  movel([-0.121105, -0.793361, -2.803748, -1.115280, 1.570796, 1.449692],accel_mss,speed_ms,0,blend_radius_m)
  movel([-0.120159, -0.793542, -2.803719, -1.115129, 1.570796, 1.450637],accel_mss,speed_ms,0,blend_radius_m)
  movel([-0.119008, -0.795086, -2.803467, -1.113836, 1.570796, 1.451789],accel_mss,speed_ms,0,blend_radius_m)
  movel([-0.118135, -0.797911, -2.803003, -1.111475, 1.570796, 1.452661],accel_mss,speed_ms,0,blend_radius_m)
  movel([-0.117601, -0.801037, -2.802486, -1.108866, 1.570796, 1.453195],accel_mss,speed_ms,0,blend_radius_m)
  movel([-0.115239, -0.796332, -2.803263, -1.112794, 1.570796, 1.455558],accel_mss,speed_ms,0,blend_radius_m)
  movel([-0.112520, -0.791566, -2.804039, -1.116785, 1.570796, 1.458276],accel_mss,speed_ms,0,blend_radius_m)
  movel([-0.109499, -0.786802, -2.804803, -1.120785, 1.570796, 1.461298],accel_mss,speed_ms,0,blend_radius_m)
  movel([-0.106241, -0.782109, -2.805544, -1.124735, 1.570796, 1.464556],accel_mss,speed_ms,0,blend_radius_m)
  movel([-0.099689, -0.772678, -2.807001, -1.132710, 1.570796, 1.471108],accel_mss,speed_ms,0,blend_radius_m)
  movel([-0.097728, -0.770078, -2.807395, -1.134915, 1.570796, 1.473068],accel_mss,speed_ms,0,blend_radius_m)
  movel([-0.095794, -0.767754, -2.807745, -1.136890, 1.570796, 1.475003],accel_mss,speed_ms,0,blend_radius_m)
  movel([-0.093954, -0.765885, -2.808024, -1.138480, 1.570796, 1.476842],accel_mss,speed_ms,0,blend_radius_m)
  movel([-0.092299, -0.764660, -2.808206, -1.139523, 1.570796, 1.478498],accel_mss,speed_ms,0,blend_radius_m)
  movel([-0.090884, -0.764292, -2.808260, -1.139836, 1.570796, 1.479912],accel_mss,speed_ms,0,blend_radius_m)
  movel([-0.089878, -0.764818, -2.808182, -1.139389, 1.570796, 1.480919],accel_mss,speed_ms,0,blend_radius_m)
  movel([-0.089251, -0.766042, -2.808000, -1.138346, 1.570796, 1.481545],accel_mss,speed_ms,0,blend_radius_m)
  movel([-0.088991, -0.767774, -2.807742, -1.136873, 1.570796, 1.481805],accel_mss,speed_ms,0,blend_radius_m)
  movel([-0.089073, -0.769817, -2.807435, -1.135137, 1.570796, 1.481724],accel_mss,speed_ms,0,blend_radius_m)
  movel([-0.089471, -0.771972, -2.807109, -1.133309, 1.570796, 1.481326],accel_mss,speed_ms,0,blend_radius_m)
  movel([-0.090165, -0.774050, -2.806792, -1.131547, 1.570796, 1.480631],accel_mss,speed_ms,0,blend_radius_m)
  movel([-0.091138, -0.775860, -2.806515, -1.130015, 1.570796, 1.479658],accel_mss,speed_ms,0,blend_radius_m)
  movel([-0.085055, -0.767504, -2.807782, -1.137103, 1.570796, 1.485742],accel_mss,speed_ms,0,blend_radius_m)
  movel([-0.081792, -0.763433, -2.808387, -1.140568, 1.570796, 1.489004],accel_mss,speed_ms,0,blend_radius_m)
  movel([-0.078396, -0.759483, -2.808967, -1.143939, 1.570796, 1.492400],accel_mss,speed_ms,0,blend_radius_m)
  movel([-0.074888, -0.755690, -2.809517, -1.147182, 1.570796, 1.495909],accel_mss,speed_ms,0,blend_radius_m)
  movel([-0.071275, -0.752094, -2.810031, -1.150264, 1.570796, 1.499521],accel_mss,speed_ms,0,blend_radius_m)
  movel([-0.067576, -0.748733, -2.810507, -1.153150, 1.570796, 1.503221],accel_mss,speed_ms,0,blend_radius_m)
  movel([-0.063806, -0.745643, -2.810939, -1.155807, 1.570796, 1.506991],accel_mss,speed_ms,0,blend_radius_m)
  movel([-0.061242, -0.744068, -2.811158, -1.157163, 1.570796, 1.509554],accel_mss,speed_ms,0,blend_radius_m)
  movel([-0.058496, -0.743084, -2.811294, -1.158011, 1.570796, 1.512301],accel_mss,speed_ms,0,blend_radius_m)
  movel([-0.057304, -0.742971, -2.811309, -1.158108, 1.570796, 1.513493],accel_mss,speed_ms,0,blend_radius_m)
  movel([-0.056360, -0.743186, -2.811280, -1.157923, 1.570796, 1.514437],accel_mss,speed_ms,0,blend_radius_m)
  movel([-0.055759, -0.743792, -2.811196, -1.157401, 1.570796, 1.515037],accel_mss,speed_ms,0,blend_radius_m)
  movel([-0.055607, -0.744852, -2.811049, -1.156488, 1.570796, 1.515190],accel_mss,speed_ms,0,blend_radius_m)
  movel([-0.055970, -0.746235, -2.810857, -1.155298, 1.570796, 1.514827],accel_mss,speed_ms,0,blend_radius_m)
  movel([-0.056714, -0.747783, -2.810640, -1.153965, 1.570796, 1.514083],accel_mss,speed_ms,0,blend_radius_m)
  movel([-0.058927, -0.751255, -2.810150, -1.150983, 1.570796, 1.511869],accel_mss,speed_ms,0,blend_radius_m)
  movel([-0.061573, -0.754500, -2.809688, -1.148201, 1.570796, 1.509223],accel_mss,speed_ms,0,blend_radius_m)
  movel([-0.064470, -0.757491, -2.809257, -1.145642, 1.570796, 1.506326],accel_mss,speed_ms,0,blend_radius_m)
  movel([-0.067437, -0.760200, -2.808862, -1.143327, 1.570796, 1.503359],accel_mss,speed_ms,0,blend_radius_m)
  movel([-0.063607, -0.758678, -2.809084, -1.144626, 1.570796, 1.507189],accel_mss,speed_ms,0,blend_radius_m)
  movel([-0.059620, -0.756697, -2.809371, -1.146320, 1.570796, 1.511176],accel_mss,speed_ms,0,blend_radius_m)
  movel([-0.055519, -0.754282, -2.809719, -1.148388, 1.570796, 1.515278],accel_mss,speed_ms,0,blend_radius_m)
  movel([-0.051338, -0.751454, -2.810122, -1.150813, 1.570796, 1.519459],accel_mss,speed_ms,0,blend_radius_m)
  movel([-0.048030, -0.748869, -2.810488, -1.153033, 1.570796, 1.522766],accel_mss,speed_ms,0,blend_radius_m)
  movel([-0.041537, -0.743272, -2.811268, -1.157849, 1.570796, 1.529259],accel_mss,speed_ms,0,blend_radius_m)
  movel([-0.038202, -0.740640, -2.811630, -1.160119, 1.570796, 1.532595],accel_mss,speed_ms,0,blend_radius_m)
  movel([-0.034400, -0.737919, -2.812001, -1.162470, 1.570796, 1.536396],accel_mss,speed_ms,0,blend_radius_m)
  movel([-0.027997, -0.733681, -2.812571, -1.166137, 1.570796, 1.542799],accel_mss,speed_ms,0,blend_radius_m)
  movel([-0.024935, -0.731926, -2.812805, -1.167658, 1.570796, 1.545861],accel_mss,speed_ms,0,blend_radius_m)
  movel([-0.022568, -0.730917, -2.812939, -1.168533, 1.570796, 1.548229],accel_mss,speed_ms,0,blend_radius_m)
  movel([-0.021784, -0.730807, -2.812954, -1.168629, 1.570796, 1.549013],accel_mss,speed_ms,0,blend_radius_m)
  movel([-0.021347, -0.731026, -2.812924, -1.168438, 1.570796, 1.549449],accel_mss,speed_ms,0,blend_radius_m)
  movel([-0.021306, -0.731611, -2.812847, -1.167931, 1.570796, 1.549490],accel_mss,speed_ms,0,blend_radius_m)
  movel([-0.021722, -0.732612, -2.812714, -1.167063, 1.570796, 1.549074],accel_mss,speed_ms,0,blend_radius_m)
  movel([-0.023301, -0.735118, -2.812379, -1.164892, 1.570796, 1.547495],accel_mss,speed_ms,0,blend_radius_m)
  movel([-0.025347, -0.737745, -2.812024, -1.162620, 1.570796, 1.545450],accel_mss,speed_ms,0,blend_radius_m)
  movel([-0.027725, -0.740428, -2.811659, -1.160302, 1.570796, 1.543072],accel_mss,speed_ms,0,blend_radius_m)
  movel([-0.030292, -0.743084, -2.811294, -1.158011, 1.570796, 1.540504],accel_mss,speed_ms,0,blend_radius_m)
  movel([-0.035478, -0.748036, -2.810605, -1.153749, 1.570796, 1.535318],accel_mss,speed_ms,0,blend_radius_m)
  movel([-0.039835, -0.752018, -2.810042, -1.150329, 1.570796, 1.530962],accel_mss,speed_ms,0,blend_radius_m)
  movel([-0.037640, -0.751618, -2.810099, -1.150672, 1.570796, 1.533156],accel_mss,speed_ms,0,blend_radius_m)
  movel([-0.035326, -0.750943, -2.810195, -1.151251, 1.570796, 1.535470],accel_mss,speed_ms,0,blend_radius_m)
  movel([-0.030418, -0.748918, -2.810481, -1.152991, 1.570796, 1.540378],accel_mss,speed_ms,0,blend_radius_m)
  movel([-0.025249, -0.746199, -2.810862, -1.155329, 1.570796, 1.545548],accel_mss,speed_ms,0,blend_radius_m)
  movel([-0.019955, -0.743049, -2.811299, -1.158041, 1.570796, 1.550841],accel_mss,speed_ms,0,blend_radius_m)
  movel([-0.015550, -0.740169, -2.811694, -1.160526, 1.570796, 1.555246],accel_mss,speed_ms,0,blend_radius_m)
  movel([-0.002182, -0.730928, -2.812937, -1.168523, 1.570796, 1.568614],accel_mss,speed_ms,0,blend_radius_m)
  movel([0.000291, -0.729638, -2.813108, -1.169643, 1.570796, 1.571087],accel_mss,speed_ms,0,blend_radius_m)
  movel([0.002219, -0.729213, -2.813164, -1.170012, 1.570796, 1.573015],accel_mss,speed_ms,0,blend_radius_m)
  movel([0.002614, -0.729532, -2.813122, -1.169735, 1.570796, 1.573410],accel_mss,speed_ms,0,blend_radius_m)
  movel([0.002432, -0.730316, -2.813018, -1.169054, 1.570796, 1.573228],accel_mss,speed_ms,0,blend_radius_m)
  movel([0.001528, -0.731648, -2.812842, -1.167899, 1.570796, 1.572325],accel_mss,speed_ms,0,blend_radius_m)
  movel([-0.000242, -0.733605, -2.812581, -1.166203, 1.570796, 1.570554],accel_mss,speed_ms,0,blend_radius_m)
  movel([-0.003204, -0.736443, -2.812200, -1.163745, 1.570796, 1.567592],accel_mss,speed_ms,0,blend_radius_m)
  movel([-0.006618, -0.739358, -2.811805, -1.161226, 1.570796, 1.564179],accel_mss,speed_ms,0,blend_radius_m)
  movel([-0.009977, -0.741812, -2.811469, -1.159108, 1.570796, 1.560819],accel_mss,speed_ms,0,blend_radius_m)
  movel([-0.011482, -0.742703, -2.811346, -1.158339, 1.570796, 1.559315],accel_mss,speed_ms,0,blend_radius_m)
  movel([-0.012779, -0.743271, -2.811268, -1.157850, 1.570796, 1.558017],accel_mss,speed_ms,0,blend_radius_m)
  movel([-0.007737, -0.743073, -2.811295, -1.158021, 1.570796, 1.563059],accel_mss,speed_ms,0,blend_radius_m)
  movel([-0.002332, -0.742171, -2.811420, -1.158799, 1.570796, 1.568464],accel_mss,speed_ms,0,blend_radius_m)
  movel([0.003362, -0.740698, -2.811622, -1.160069, 1.570796, 1.574158],accel_mss,speed_ms,0,blend_radius_m)
  movel([0.009278, -0.738793, -2.811882, -1.161714, 1.570796, 1.580074],accel_mss,speed_ms,0,blend_radius_m)
  movel([0.021466, -0.734216, -2.812500, -1.165673, 1.570796, 1.592262],accel_mss,speed_ms,0,blend_radius_m)
  movel([0.033600, -0.729546, -2.813120, -1.169723, 1.570796, 1.604396],accel_mss,speed_ms,0,blend_radius_m)
  movel([0.035605, -0.729117, -2.813177, -1.170096, 1.570796, 1.606402],accel_mss,speed_ms,0,blend_radius_m)
  movel([0.036255, -0.729398, -2.813140, -1.169851, 1.570796, 1.607051],accel_mss,speed_ms,0,blend_radius_m)
  movel([0.036422, -0.730219, -2.813031, -1.169139, 1.570796, 1.607218],accel_mss,speed_ms,0,blend_radius_m)
  movel([0.036036, -0.731427, -2.812871, -1.168090, 1.570796, 1.606833],accel_mss,speed_ms,0,blend_radius_m)
  movel([0.034004, -0.734771, -2.812425, -1.165193, 1.570796, 1.604800],accel_mss,speed_ms,0,blend_radius_m)
  movel([0.032557, -0.736690, -2.812167, -1.163532, 1.570796, 1.603354],accel_mss,speed_ms,0,blend_radius_m)
  movel([0.029315, -0.740256, -2.811682, -1.160451, 1.570796, 1.600111],accel_mss,speed_ms,0,blend_radius_m)
  movel([0.025758, -0.743429, -2.811246, -1.157714, 1.570796, 1.596555],accel_mss,speed_ms,0,blend_radius_m)
  movel([0.022037, -0.746209, -2.810860, -1.155320, 1.570796, 1.592834],accel_mss,speed_ms,0,blend_radius_m)
  movel([0.018315, -0.748574, -2.810529, -1.153286, 1.570796, 1.589112],accel_mss,speed_ms,0,blend_radius_m)
  movel([0.014745, -0.750516, -2.810255, -1.151618, 1.570796, 1.585541],accel_mss,speed_ms,0,blend_radius_m)
  movel([0.011481, -0.752014, -2.810043, -1.150332, 1.570796, 1.582277],accel_mss,speed_ms,0,blend_radius_m)
  movel([0.008687, -0.753044, -2.809896, -1.149449, 1.570796, 1.579483],accel_mss,speed_ms,0,blend_radius_m)
  movel([0.008653, -0.753899, -2.809774, -1.148717, 1.570796, 1.579449],accel_mss,speed_ms,0,blend_radius_m)
  movel([0.009139, -0.754307, -2.809715, -1.148367, 1.570796, 1.579935],accel_mss,speed_ms,0,blend_radius_m)
  movel([0.010647, -0.754705, -2.809658, -1.148026, 1.570796, 1.581444],accel_mss,speed_ms,0,blend_radius_m)
  movel([0.012360, -0.754771, -2.809649, -1.147969, 1.570796, 1.583157],accel_mss,speed_ms,0,blend_radius_m)
  movel([0.016128, -0.754316, -2.809714, -1.148359, 1.570796, 1.586925],accel_mss,speed_ms,0,blend_radius_m)
  movel([0.022850, -0.753072, -2.809892, -1.149425, 1.570796, 1.593647],accel_mss,speed_ms,0,blend_radius_m)
  movel([0.029687, -0.751537, -2.810110, -1.150742, 1.570796, 1.600483],accel_mss,speed_ms,0,blend_radius_m)
  movel([0.043712, -0.747708, -2.810651, -1.154030, 1.570796, 1.614508],accel_mss,speed_ms,0,blend_radius_m)
  movel([0.047601, -0.746731, -2.810787, -1.154870, 1.570796, 1.618397],accel_mss,speed_ms,0,blend_radius_m)
  movel([0.050057, -0.746348, -2.810841, -1.155200, 1.570796, 1.620854],accel_mss,speed_ms,0,blend_radius_m)
  movel([0.052405, -0.746275, -2.810851, -1.155263, 1.570796, 1.623201],accel_mss,speed_ms,0,blend_radius_m)
  movel([0.054288, -0.746698, -2.810792, -1.154899, 1.570796, 1.625084],accel_mss,speed_ms,0,blend_radius_m)
  movel([0.055366, -0.747783, -2.810640, -1.153965, 1.570796, 1.626162],accel_mss,speed_ms,0,blend_radius_m)
  movel([0.055503, -0.748623, -2.810522, -1.153244, 1.570796, 1.626300],accel_mss,speed_ms,0,blend_radius_m)
  movel([0.055317, -0.749691, -2.810372, -1.152326, 1.570796, 1.626113],accel_mss,speed_ms,0,blend_radius_m)
  movel([0.054755, -0.751016, -2.810184, -1.151188, 1.570796, 1.625552],accel_mss,speed_ms,0,blend_radius_m)
  movel([0.053791, -0.752605, -2.809958, -1.149825, 1.570796, 1.624588],accel_mss,speed_ms,0,blend_radius_m)
  movel([0.052380, -0.754061, -2.809750, -1.148578, 1.570796, 1.623176],accel_mss,speed_ms,0,blend_radius_m)
  movel([0.050460, -0.755437, -2.809553, -1.147399, 1.570796, 1.621256],accel_mss,speed_ms,0,blend_radius_m)
  movel([0.040183, -0.761646, -2.808651, -1.142093, 1.570796, 1.610979],accel_mss,speed_ms,0,blend_radius_m)
  movel([0.036738, -0.763274, -2.808411, -1.140704, 1.570796, 1.607535],accel_mss,speed_ms,0,blend_radius_m)
  movel([0.035260, -0.763727, -2.808344, -1.140318, 1.570796, 1.606056],accel_mss,speed_ms,0,blend_radius_m)
  movel([0.034042, -0.763830, -2.808329, -1.140230, 1.570796, 1.604838],accel_mss,speed_ms,0,blend_radius_m)
  movel([0.039097, -0.765388, -2.808098, -1.138903, 1.570796, 1.609893],accel_mss,speed_ms,0,blend_radius_m)
  movel([0.044720, -0.766036, -2.808001, -1.138351, 1.570796, 1.615516],accel_mss,speed_ms,0,blend_radius_m)
  movel([0.050778, -0.765942, -2.808015, -1.138432, 1.570796, 1.621574],accel_mss,speed_ms,0,blend_radius_m)
  movel([0.057144, -0.765260, -2.808117, -1.139012, 1.570796, 1.627940],accel_mss,speed_ms,0,blend_radius_m)
  movel([0.062648, -0.763858, -2.808325, -1.140207, 1.570796, 1.633444],accel_mss,speed_ms,0,blend_radius_m)
  movel([0.070534, -0.762014, -2.808596, -1.141778, 1.570796, 1.641330],accel_mss,speed_ms,0,blend_radius_m)
  movel([0.074102, -0.761631, -2.808653, -1.142105, 1.570796, 1.644899],accel_mss,speed_ms,0,blend_radius_m)
  movel([0.076754, -0.761962, -2.808604, -1.141823, 1.570796, 1.647550],accel_mss,speed_ms,0,blend_radius_m)
  movel([0.077577, -0.762479, -2.808528, -1.141382, 1.570796, 1.648374],accel_mss,speed_ms,0,blend_radius_m)
  movel([0.077981, -0.763272, -2.808411, -1.140706, 1.570796, 1.648777],accel_mss,speed_ms,0,blend_radius_m)
  movel([0.077904, -0.764377, -2.808248, -1.139764, 1.570796, 1.648701],accel_mss,speed_ms,0,blend_radius_m)
  movel([0.077296, -0.765814, -2.808034, -1.138540, 1.570796, 1.648093],accel_mss,speed_ms,0,blend_radius_m)
  movel([0.076368, -0.767285, -2.807815, -1.137289, 1.570796, 1.647164],accel_mss,speed_ms,0,blend_radius_m)
  movel([0.075295, -0.768687, -2.807605, -1.136097, 1.570796, 1.646091],accel_mss,speed_ms,0,blend_radius_m)
  movel([0.072924, -0.771293, -2.807212, -1.133884, 1.570796, 1.643720],accel_mss,speed_ms,0,blend_radius_m)
  movel([0.070302, -0.773862, -2.806821, -1.131706, 1.570796, 1.641099],accel_mss,speed_ms,0,blend_radius_m)
  movel([0.064988, -0.778418, -2.806120, -1.127851, 1.570796, 1.635784],accel_mss,speed_ms,0,blend_radius_m)
  movel([0.062326, -0.780386, -2.805814, -1.126189, 1.570796, 1.633122],accel_mss,speed_ms,0,blend_radius_m)
  movel([0.067181, -0.779786, -2.805907, -1.126695, 1.570796, 1.637977],accel_mss,speed_ms,0,blend_radius_m)
  movel([0.072189, -0.778807, -2.806060, -1.127523, 1.570796, 1.642985],accel_mss,speed_ms,0,blend_radius_m)
  movel([0.077338, -0.777493, -2.806263, -1.128633, 1.570796, 1.648134],accel_mss,speed_ms,0,blend_radius_m)
  movel([0.082615, -0.775877, -2.806512, -1.130000, 1.570796, 1.653412],accel_mss,speed_ms,0,blend_radius_m)
  movel([0.093490, -0.771912, -2.807118, -1.133359, 1.570796, 1.664286],accel_mss,speed_ms,0,blend_radius_m)
  movel([0.104701, -0.767216, -2.807825, -1.137348, 1.570796, 1.675497],accel_mss,speed_ms,0,blend_radius_m)
  movel([0.107639, -0.766300, -2.807962, -1.138127, 1.570796, 1.678435],accel_mss,speed_ms,0,blend_radius_m)
  movel([0.108683, -0.766493, -2.807933, -1.137963, 1.570796, 1.679480],accel_mss,speed_ms,0,blend_radius_m)
  movel([0.109107, -0.767448, -2.807791, -1.137151, 1.570796, 1.679903],accel_mss,speed_ms,0,blend_radius_m)
  movel([0.108974, -0.768426, -2.807644, -1.136319, 1.570796, 1.679770],accel_mss,speed_ms,0,blend_radius_m)
  movel([0.108569, -0.769523, -2.807479, -1.135387, 1.570796, 1.679365],accel_mss,speed_ms,0,blend_radius_m)
  movel([0.107060, -0.772017, -2.807102, -1.133270, 1.570796, 1.677856],accel_mss,speed_ms,0,blend_radius_m)
  movel([0.104857, -0.774737, -2.806687, -1.130965, 1.570796, 1.675653],accel_mss,speed_ms,0,blend_radius_m)
  movel([0.102226, -0.777515, -2.806260, -1.128615, 1.570796, 1.673022],accel_mss,speed_ms,0,blend_radius_m)
  movel([0.096762, -0.782520, -2.805480, -1.124390, 1.570796, 1.667558],accel_mss,speed_ms,0,blend_radius_m)
  movel([0.092780, -0.785621, -2.804990, -1.121778, 1.570796, 1.663577],accel_mss,speed_ms,0,blend_radius_m)
  movel([0.095018, -0.784942, -2.805098, -1.122349, 1.570796, 1.665815],accel_mss,speed_ms,0,blend_radius_m)
  movel([0.097342, -0.784002, -2.805247, -1.123140, 1.570796, 1.668138],accel_mss,speed_ms,0,blend_radius_m)
  movel([0.102193, -0.781425, -2.805652, -1.125313, 1.570796, 1.672990],accel_mss,speed_ms,0,blend_radius_m)
  movel([0.107238, -0.777995, -2.806185, -1.128209, 1.570796, 1.678035],accel_mss,speed_ms,0,blend_radius_m)
  movel([0.112383, -0.773843, -2.806824, -1.131722, 1.570796, 1.683179],accel_mss,speed_ms,0,blend_radius_m)
  movel([0.117534, -0.769067, -2.807548, -1.135774, 1.570796, 1.688330],accel_mss,speed_ms,0,blend_radius_m)
  movel([0.122590, -0.763799, -2.808333, -1.140256, 1.570796, 1.693387],accel_mss,speed_ms,0,blend_radius_m)
  movel([0.127452, -0.758145, -2.809162, -1.145082, 1.570796, 1.698249],accel_mss,speed_ms,0,blend_radius_m)
  movel([0.132018, -0.752235, -2.810011, -1.150143, 1.570796, 1.702814],accel_mss,speed_ms,0,blend_radius_m)
  movel([0.134037, -0.749592, -2.810386, -1.152411, 1.570796, 1.704834],accel_mss,speed_ms,0,blend_radius_m)
  movel([0.135120, -0.748440, -2.810548, -1.153401, 1.570796, 1.705916],accel_mss,speed_ms,0,blend_radius_m)
  movel([0.136237, -0.747552, -2.810672, -1.154164, 1.570796, 1.707033],accel_mss,speed_ms,0,blend_radius_m)
  movel([0.137379, -0.747065, -2.810741, -1.154583, 1.570796, 1.708175],accel_mss,speed_ms,0,blend_radius_m)
  movel([0.138333, -0.747027, -2.810746, -1.154616, 1.570796, 1.709129],accel_mss,speed_ms,0,blend_radius_m)
  movel([0.139345, -0.747698, -2.810652, -1.154039, 1.570796, 1.710141],accel_mss,speed_ms,0,blend_radius_m)
  movel([0.139829, -0.749137, -2.810450, -1.152802, 1.570796, 1.710625],accel_mss,speed_ms,0,blend_radius_m)
  movel([0.139879, -0.751150, -2.810165, -1.151074, 1.570796, 1.710675],accel_mss,speed_ms,0,blend_radius_m)
  movel([0.139591, -0.753557, -2.809823, -1.149009, 1.570796, 1.710387],accel_mss,speed_ms,0,blend_radius_m)
  movel([0.138373, -0.758783, -2.809069, -1.144537, 1.570796, 1.709169],accel_mss,speed_ms,0,blend_radius_m)
  movel([0.136926, -0.763333, -2.808402, -1.140654, 1.570796, 1.707723],accel_mss,speed_ms,0,blend_radius_m)
  movel([0.140852, -0.757577, -2.809244, -1.145568, 1.570796, 1.711648],accel_mss,speed_ms,0,blend_radius_m)
  movel([0.144402, -0.751708, -2.810086, -1.150595, 1.570796, 1.715198],accel_mss,speed_ms,0,blend_radius_m)
  movel([0.147549, -0.745784, -2.810919, -1.155685, 1.570796, 1.718345],accel_mss,speed_ms,0,blend_radius_m)
  movel([0.150273, -0.739888, -2.811733, -1.160768, 1.570796, 1.721070],accel_mss,speed_ms,0,blend_radius_m)
  movel([0.152533, -0.734096, -2.812516, -1.165777, 1.570796, 1.723330],accel_mss,speed_ms,0,blend_radius_m)
  movel([0.154318, -0.728473, -2.813261, -1.170655, 1.570796, 1.725114],accel_mss,speed_ms,0,blend_radius_m)
  movel([0.155580, -0.723118, -2.813958, -1.175313, 1.570796, 1.726376],accel_mss,speed_ms,0,blend_radius_m)
  movel([0.156297, -0.718102, -2.814598, -1.179688, 1.570796, 1.727094],accel_mss,speed_ms,0,blend_radius_m)
  movel([0.156402, -0.711752, -2.815393, -1.185243, 1.570796, 1.727198],accel_mss,speed_ms,0,blend_radius_m)
  movel([0.156716, -0.708235, -2.815826, -1.188328, 1.570796, 1.727512],accel_mss,speed_ms,0,blend_radius_m)
  movel([0.157110, -0.706436, -2.816045, -1.189908, 1.570796, 1.727906],accel_mss,speed_ms,0,blend_radius_m)
  movel([0.157721, -0.704629, -2.816264, -1.191496, 1.570796, 1.728517],accel_mss,speed_ms,0,blend_radius_m)
  movel([0.159157, -0.701655, -2.816621, -1.194114, 1.570796, 1.729953],accel_mss,speed_ms,0,blend_radius_m)
  movel([0.160486, -0.699829, -2.816838, -1.195722, 1.570796, 1.731283],accel_mss,speed_ms,0,blend_radius_m)
  movel([0.161725, -0.698910, -2.816946, -1.196533, 1.570796, 1.732521],accel_mss,speed_ms,0,blend_radius_m)
  movel([0.162880, -0.698652, -2.816977, -1.196760, 1.570796, 1.733676],accel_mss,speed_ms,0,blend_radius_m)
  movel([0.165920, -0.699423, -2.816886, -1.196081, 1.570796, 1.736716],accel_mss,speed_ms,0,blend_radius_m)
  movel([0.166833, -0.699369, -2.816892, -1.196128, 1.570796, 1.737629],accel_mss,speed_ms,0,blend_radius_m)
  movel([0.168876, -0.694954, -2.817410, -1.200024, 1.570796, 1.739672],accel_mss,speed_ms,0,blend_radius_m)
  movel([0.170617, -0.690579, -2.817915, -1.203895, 1.570796, 1.741413],accel_mss,speed_ms,0,blend_radius_m)
  movel([0.172069, -0.686262, -2.818406, -1.207721, 1.570796, 1.742866],accel_mss,speed_ms,0,blend_radius_m)
  movel([0.173248, -0.682014, -2.818880, -1.211495, 1.570796, 1.744044],accel_mss,speed_ms,0,blend_radius_m)
  movel([0.174153, -0.677863, -2.819337, -1.215189, 1.570796, 1.744950],accel_mss,speed_ms,0,blend_radius_m)
  movel([0.174801, -0.673819, -2.819775, -1.218796, 1.570796, 1.745598],accel_mss,speed_ms,0,blend_radius_m)
  movel([0.175391, -0.666110, -2.820590, -1.225689, 1.570796, 1.746188],accel_mss,speed_ms,0,blend_radius_m)
  movel([0.175103, -0.659042, -2.821316, -1.232031, 1.570796, 1.745899],accel_mss,speed_ms,0,blend_radius_m)
  movel([0.174059, -0.652731, -2.821947, -1.237712, 1.570796, 1.744855],accel_mss,speed_ms,0,blend_radius_m)
  movel([0.172351, -0.647325, -2.822474, -1.242590, 1.570796, 1.743147],accel_mss,speed_ms,0,blend_radius_m)
  movel([0.170116, -0.642932, -2.822894, -1.246563, 1.570796, 1.740912],accel_mss,speed_ms,0,blend_radius_m)
  speed_ms = 0.005
  movel([0.170116, -0.636489, -2.816133, -1.259767, 1.570796, 1.740912],accel_mss,speed_ms,0,blend_radius_m)
  speed_ms = 0.040
  movel([0.138700, -0.661451, -2.813652, -1.237286, 1.570796, 1.709497],accel_mss,speed_ms,0,blend_radius_m)
  speed_ms = 0.005
  movel([0.138700, -0.668285, -2.820362, -1.223742, 1.570796, 1.709497],accel_mss,speed_ms,0,blend_radius_m)
  speed_ms = 0.025
  movel([0.136102, -0.667914, -2.820401, -1.224074, 1.570796, 1.706899],accel_mss,speed_ms,0,blend_radius_m)
  movel([0.133054, -0.668449, -2.820345, -1.223595, 1.570796, 1.703850],accel_mss,speed_ms,0,blend_radius_m)
  movel([0.129644, -0.669757, -2.820207, -1.222425, 1.570796, 1.700441],accel_mss,speed_ms,0,blend_radius_m)
  movel([0.125976, -0.671690, -2.820002, -1.220697, 1.570796, 1.696772],accel_mss,speed_ms,0,blend_radius_m)
  movel([0.122143, -0.674109, -2.819743, -1.218536, 1.570796, 1.692939],accel_mss,speed_ms,0,blend_radius_m)
  movel([0.118234, -0.676875, -2.819444, -1.216069, 1.570796, 1.689030],accel_mss,speed_ms,0,blend_radius_m)
  movel([0.110564, -0.682887, -2.818784, -1.210719, 1.570796, 1.681360],accel_mss,speed_ms,0,blend_radius_m)
  speed_ms = 0.005
  movel([0.110564, -0.675837, -2.812104, -1.224448, 1.570796, 1.681360],accel_mss,speed_ms,0,blend_radius_m)
  speed_ms = 0.040
  movel([0.120496, -0.667301, -2.813033, -1.232055, 1.570796, 1.691293],accel_mss,speed_ms,0,blend_radius_m)
  speed_ms = 0.005
  movel([0.120496, -0.674223, -2.819731, -1.218435, 1.570796, 1.691293],accel_mss,speed_ms,0,blend_radius_m)
  speed_ms = 0.025
  movel([0.122110, -0.669388, -2.820246, -1.222755, 1.570796, 1.692907],accel_mss,speed_ms,0,blend_radius_m)
  movel([0.123299, -0.664893, -2.820716, -1.226780, 1.570796, 1.694095],accel_mss,speed_ms,0,blend_radius_m)
  movel([0.124068, -0.660732, -2.821144, -1.230512, 1.570796, 1.694864],accel_mss,speed_ms,0,blend_radius_m)
  movel([0.124435, -0.656891, -2.821533, -1.233966, 1.570796, 1.695231],accel_mss,speed_ms,0,blend_radius_m)
  movel([0.124423, -0.653347, -2.821886, -1.237156, 1.570796, 1.695219],accel_mss,speed_ms,0,blend_radius_m)
  movel([0.124046, -0.650090, -2.822206, -1.240093, 1.570796, 1.694842],accel_mss,speed_ms,0,blend_radius_m)
  movel([0.123323, -0.647102, -2.822495, -1.242791, 1.570796, 1.694119],accel_mss,speed_ms,0,blend_radius_m)
  movel([0.122274, -0.644366, -2.822758, -1.245265, 1.570796, 1.693071],accel_mss,speed_ms,0,blend_radius_m)
  movel([0.118229, -0.637367, -2.823415, -1.251608, 1.570796, 1.689025],accel_mss,speed_ms,0,blend_radius_m)
  movel([0.116481, -0.633814, -2.823740, -1.254834, 1.570796, 1.687277],accel_mss,speed_ms,0,blend_radius_m)
  movel([0.115290, -0.629199, -2.824156, -1.259034, 1.570796, 1.686086],accel_mss,speed_ms,0,blend_radius_m)
  movel([0.114590, -0.622661, -2.824731, -1.264997, 1.570796, 1.685386],accel_mss,speed_ms,0,blend_radius_m)
  movel([0.114549, -0.615508, -2.825341, -1.271541, 1.570796, 1.685345],accel_mss,speed_ms,0,blend_radius_m)
  movel([0.115398, -0.607615, -2.825990, -1.278783, 1.570796, 1.686195],accel_mss,speed_ms,0,blend_radius_m)
  movel([0.116229, -0.603351, -2.826331, -1.282706, 1.570796, 1.687025],accel_mss,speed_ms,0,blend_radius_m)
  movel([0.117376, -0.598855, -2.826683, -1.286851, 1.570796, 1.688172],accel_mss,speed_ms,0,blend_radius_m)
  movel([0.119840, -0.591525, -2.827240, -1.293623, 1.570796, 1.690636],accel_mss,speed_ms,0,blend_radius_m)
  movel([0.123098, -0.583987, -2.827792, -1.300610, 1.570796, 1.693894],accel_mss,speed_ms,0,blend_radius_m)
  movel([0.127112, -0.576293, -2.828334, -1.307763, 1.570796, 1.697908],accel_mss,speed_ms,0,blend_radius_m)
  movel([0.131842, -0.568506, -2.828859, -1.315023, 1.570796, 1.702638],accel_mss,speed_ms,0,blend_radius_m)
  movel([0.137234, -0.560707, -2.829363, -1.322319, 1.570796, 1.708030],accel_mss,speed_ms,0,blend_radius_m)
  movel([0.143247, -0.552962, -2.829842, -1.329585, 1.570796, 1.714044],accel_mss,speed_ms,0,blend_radius_m)
  movel([0.149829, -0.545343, -2.830291, -1.336755, 1.570796, 1.720625],accel_mss,speed_ms,0,blend_radius_m)
  movel([0.156913, -0.537942, -2.830707, -1.343739, 1.570796, 1.727709],accel_mss,speed_ms,0,blend_radius_m)
  movel([0.162439, -0.532674, -2.830992, -1.348723, 1.570796, 1.733235],accel_mss,speed_ms,0,blend_radius_m)
  movel([0.168059, -0.527738, -2.831250, -1.353401, 1.570796, 1.738855],accel_mss,speed_ms,0,blend_radius_m)
  movel([0.173713, -0.523179, -2.831480, -1.357730, 1.570796, 1.744510],accel_mss,speed_ms,0,blend_radius_m)
  movel([0.179359, -0.519012, -2.831684, -1.361692, 1.570796, 1.750155],accel_mss,speed_ms,0,blend_radius_m)
  movel([0.184932, -0.515296, -2.831861, -1.365232, 1.570796, 1.755728],accel_mss,speed_ms,0,blend_radius_m)
  movel([0.190379, -0.512056, -2.832011, -1.368322, 1.570796, 1.761175],accel_mss,speed_ms,0,blend_radius_m)
  movel([0.195640, -0.509329, -2.832135, -1.370925, 1.570796, 1.766437],accel_mss,speed_ms,0,blend_radius_m)
  movel([0.200660, -0.507152, -2.832232, -1.373005, 1.570796, 1.771456],accel_mss,speed_ms,0,blend_radius_m)
  movel([0.205378, -0.505561, -2.832301, -1.374527, 1.570796, 1.776175],accel_mss,speed_ms,0,blend_radius_m)
  movel([0.209750, -0.504576, -2.832344, -1.375469, 1.570796, 1.780546],accel_mss,speed_ms,0,blend_radius_m)
  movel([0.213716, -0.504236, -2.832359, -1.375794, 1.570796, 1.784512],accel_mss,speed_ms,0,blend_radius_m)
  movel([0.217226, -0.504564, -2.832345, -1.375480, 1.570796, 1.788023],accel_mss,speed_ms,0,blend_radius_m)
  movel([0.220235, -0.505581, -2.832300, -1.374508, 1.570796, 1.791031],accel_mss,speed_ms,0,blend_radius_m)
  movel([0.222682, -0.507322, -2.832224, -1.372843, 1.570796, 1.793478],accel_mss,speed_ms,0,blend_radius_m)
  movel([0.224532, -0.509791, -2.832114, -1.370484, 1.570796, 1.795329],accel_mss,speed_ms,0,blend_radius_m)
  movel([0.225745, -0.513014, -2.831967, -1.367408, 1.570796, 1.796541],accel_mss,speed_ms,0,blend_radius_m)
  movel([0.226531, -0.518024, -2.831732, -1.362634, 1.570796, 1.797328],accel_mss,speed_ms,0,blend_radius_m)
  movel([0.226728, -0.523593, -2.831459, -1.357336, 1.570796, 1.797524],accel_mss,speed_ms,0,blend_radius_m)
  movel([0.226455, -0.529591, -2.831154, -1.351644, 1.570796, 1.797251],accel_mss,speed_ms,0,blend_radius_m)
  movel([0.225856, -0.535853, -2.830821, -1.345714, 1.570796, 1.796653],accel_mss,speed_ms,0,blend_radius_m)
  movel([0.223911, -0.549926, -2.830023, -1.332440, 1.570796, 1.794707],accel_mss,speed_ms,0,blend_radius_m)
  movel([0.221348, -0.564429, -2.829125, -1.318835, 1.570796, 1.792145],accel_mss,speed_ms,0,blend_radius_m)
  movel([0.218336, -0.579212, -2.828131, -1.305046, 1.570796, 1.789132],accel_mss,speed_ms,0,blend_radius_m)
  movel([0.215033, -0.594113, -2.827046, -1.291230, 1.570796, 1.785830],accel_mss,speed_ms,0,blend_radius_m)
  movel([0.201838, -0.652335, -2.821986, -1.238068, 1.570796, 1.772635],accel_mss,speed_ms,0,blend_radius_m)
  movel([0.196552, -0.679655, -2.819141, -1.213593, 1.570796, 1.767348],accel_mss,speed_ms,0,blend_radius_m)
  movel([0.194383, -0.692825, -2.817657, -1.201907, 1.570796, 1.765179],accel_mss,speed_ms,0,blend_radius_m)
  movel([0.192649, -0.705556, -2.816152, -1.190681, 1.570796, 1.763445],accel_mss,speed_ms,0,blend_radius_m)
  movel([0.191422, -0.717796, -2.814637, -1.179956, 1.570796, 1.762219],accel_mss,speed_ms,0,blend_radius_m)
  movel([0.190783, -0.729475, -2.813129, -1.169785, 1.570796, 1.761579],accel_mss,speed_ms,0,blend_radius_m)
  movel([0.190794, -0.740548, -2.811642, -1.160199, 1.570796, 1.761590],accel_mss,speed_ms,0,blend_radius_m)
  movel([0.191537, -0.750956, -2.810193, -1.151240, 1.570796, 1.762333],accel_mss,speed_ms,0,blend_radius_m)
  movel([0.192118, -0.754746, -2.809652, -1.147991, 1.570796, 1.762914],accel_mss,speed_ms,0,blend_radius_m)
  movel([0.193186, -0.758057, -2.809174, -1.145158, 1.570796, 1.763982],accel_mss,speed_ms,0,blend_radius_m)
  movel([0.194999, -0.760444, -2.808827, -1.143118, 1.570796, 1.765795],accel_mss,speed_ms,0,blend_radius_m)
  movel([0.196267, -0.761152, -2.808723, -1.142514, 1.570796, 1.767064],accel_mss,speed_ms,0,blend_radius_m)
  movel([0.197826, -0.761455, -2.808679, -1.142255, 1.570796, 1.768623],accel_mss,speed_ms,0,blend_radius_m)
  speed_ms = 0.005
  movel([0.197826, -0.753361, -2.802191, -1.156837, 1.570796, 1.768623],accel_mss,speed_ms,0,blend_radius_m)
  speed_ms = 0.040
  movel([0.166317, -0.715093, -2.807424, -1.189872, 1.570796, 1.737113],accel_mss,speed_ms,0,blend_radius_m)
  speed_ms = 0.005
  movel([0.166317, -0.722698, -2.814012, -1.175679, 1.570796, 1.737113],accel_mss,speed_ms,0,blend_radius_m)
  speed_ms = 0.025
  movel([0.165098, -0.724655, -2.813759, -1.173975, 1.570796, 1.735894],accel_mss,speed_ms,0,blend_radius_m)
  movel([0.164169, -0.726654, -2.813499, -1.172236, 1.570796, 1.734965],accel_mss,speed_ms,0,blend_radius_m)
  movel([0.163511, -0.728662, -2.813236, -1.170490, 1.570796, 1.734307],accel_mss,speed_ms,0,blend_radius_m)
  movel([0.163074, -0.730695, -2.812968, -1.168725, 1.570796, 1.733870],accel_mss,speed_ms,0,blend_radius_m)
  movel([0.162764, -0.734758, -2.812427, -1.165204, 1.570796, 1.733560],accel_mss,speed_ms,0,blend_radius_m)
  movel([0.162975, -0.738769, -2.811885, -1.161734, 1.570796, 1.733771],accel_mss,speed_ms,0,blend_radius_m)
  movel([0.164204, -0.749737, -2.810365, -1.152287, 1.570796, 1.735001],accel_mss,speed_ms,0,blend_radius_m)
  movel([0.163980, -0.752776, -2.809934, -1.149679, 1.570796, 1.734776],accel_mss,speed_ms,0,blend_radius_m)
  movel([0.163462, -0.754289, -2.809718, -1.148382, 1.570796, 1.734258],accel_mss,speed_ms,0,blend_radius_m)
  movel([0.162572, -0.755584, -2.809532, -1.147273, 1.570796, 1.733369],accel_mss,speed_ms,0,blend_radius_m)
  movel([0.161731, -0.756362, -2.809420, -1.146608, 1.570796, 1.732527],accel_mss,speed_ms,0,blend_radius_m)
  movel([0.160936, -0.756679, -2.809374, -1.146336, 1.570796, 1.731733],accel_mss,speed_ms,0,blend_radius_m)
  movel([0.160186, -0.756603, -2.809385, -1.146401, 1.570796, 1.730982],accel_mss,speed_ms,0,blend_radius_m)
  movel([0.158834, -0.755474, -2.809548, -1.147367, 1.570796, 1.729630],accel_mss,speed_ms,0,blend_radius_m)
  movel([0.157687, -0.753438, -2.809840, -1.149111, 1.570796, 1.728483],accel_mss,speed_ms,0,blend_radius_m)
  movel([0.156071, -0.748461, -2.810545, -1.153383, 1.570796, 1.726867],accel_mss,speed_ms,0,blend_radius_m)
  movel([0.155517, -0.745304, -2.810986, -1.156098, 1.570796, 1.726314],accel_mss,speed_ms,0,blend_radius_m)
  movel([0.153840, -0.750973, -2.810190, -1.151225, 1.570796, 1.724636],accel_mss,speed_ms,0,blend_radius_m)
  movel([0.152864, -0.756252, -2.809436, -1.146702, 1.570796, 1.723661],accel_mss,speed_ms,0,blend_radius_m)
  movel([0.152485, -0.761172, -2.808720, -1.142497, 1.570796, 1.723281],accel_mss,speed_ms,0,blend_radius_m)
  movel([0.152612, -0.765738, -2.808046, -1.138605, 1.570796, 1.723409],accel_mss,speed_ms,0,blend_radius_m)
  movel([0.153139, -0.769987, -2.807409, -1.134993, 1.570796, 1.723935],accel_mss,speed_ms,0,blend_radius_m)
  movel([0.153986, -0.773916, -2.806813, -1.131660, 1.570796, 1.724782],accel_mss,speed_ms,0,blend_radius_m)
  movel([0.156246, -0.780895, -2.805734, -1.125760, 1.570796, 1.727042],accel_mss,speed_ms,0,blend_radius_m)
  movel([0.156304, -0.782559, -2.805474, -1.124357, 1.570796, 1.727100],accel_mss,speed_ms,0,blend_radius_m)
  movel([0.155931, -0.783505, -2.805325, -1.123559, 1.570796, 1.726728],accel_mss,speed_ms,0,blend_radius_m)
  movel([0.155223, -0.784307, -2.805198, -1.122883, 1.570796, 1.726019],accel_mss,speed_ms,0,blend_radius_m)
  movel([0.154317, -0.784694, -2.805137, -1.122558, 1.570796, 1.725113],accel_mss,speed_ms,0,blend_radius_m)
  movel([0.152367, -0.784864, -2.805110, -1.122415, 1.570796, 1.723163],accel_mss,speed_ms,0,blend_radius_m)
  movel([0.150735, -0.784523, -2.805164, -1.122702, 1.570796, 1.721532],accel_mss,speed_ms,0,blend_radius_m)
  movel([0.149384, -0.783748, -2.805287, -1.123355, 1.570796, 1.720180],accel_mss,speed_ms,0,blend_radius_m)
  movel([0.148290, -0.782592, -2.805469, -1.124329, 1.570796, 1.719086],accel_mss,speed_ms,0,blend_radius_m)
  movel([0.146758, -0.779427, -2.805963, -1.126999, 1.570796, 1.717554],accel_mss,speed_ms,0,blend_radius_m)
  movel([0.145914, -0.775561, -2.806561, -1.130267, 1.570796, 1.716710],accel_mss,speed_ms,0,blend_radius_m)
  movel([0.145148, -0.784445, -2.805177, -1.122768, 1.570796, 1.715944],accel_mss,speed_ms,0,blend_radius_m)
  movel([0.145196, -0.788510, -2.804530, -1.119349, 1.570796, 1.715993],accel_mss,speed_ms,0,blend_radius_m)
  movel([0.145776, -0.792154, -2.803944, -1.116291, 1.570796, 1.716573],accel_mss,speed_ms,0,blend_radius_m)
  movel([0.146955, -0.794701, -2.803530, -1.114158, 1.570796, 1.717752],accel_mss,speed_ms,0,blend_radius_m)
  movel([0.150125, -0.798602, -2.802889, -1.110898, 1.570796, 1.720921],accel_mss,speed_ms,0,blend_radius_m)
  movel([0.151210, -0.801126, -2.802471, -1.108792, 1.570796, 1.722006],accel_mss,speed_ms,0,blend_radius_m)
  movel([0.151294, -0.801757, -2.802366, -1.108266, 1.570796, 1.722090],accel_mss,speed_ms,0,blend_radius_m)
  movel([0.151105, -0.802551, -2.802233, -1.107605, 1.570796, 1.721902],accel_mss,speed_ms,0,blend_radius_m)
  movel([0.150490, -0.803397, -2.802092, -1.106900, 1.570796, 1.721287],accel_mss,speed_ms,0,blend_radius_m)
  movel([0.149467, -0.804207, -2.801956, -1.106226, 1.570796, 1.720263],accel_mss,speed_ms,0,blend_radius_m)
  movel([0.146733, -0.805659, -2.801711, -1.105019, 1.570796, 1.717529],accel_mss,speed_ms,0,blend_radius_m)
  movel([0.142223, -0.807339, -2.801427, -1.103623, 1.570796, 1.713020],accel_mss,speed_ms,0,blend_radius_m)
  movel([0.142758, -0.809563, -2.801048, -1.101778, 1.570796, 1.713554],accel_mss,speed_ms,0,blend_radius_m)
  movel([0.143619, -0.811943, -2.800640, -1.099805, 1.570796, 1.714415],accel_mss,speed_ms,0,blend_radius_m)
  movel([0.144902, -0.814307, -2.800232, -1.097850, 1.570796, 1.715698],accel_mss,speed_ms,0,blend_radius_m)
  movel([0.146705, -0.816485, -2.799853, -1.096051, 1.570796, 1.717501],accel_mss,speed_ms,0,blend_radius_m)
  movel([0.152042, -0.818606, -2.799482, -1.094301, 1.570796, 1.722838],accel_mss,speed_ms,0,blend_radius_m)
  movel([0.154980, -0.819950, -2.799245, -1.093193, 1.570796, 1.725776],accel_mss,speed_ms,0,blend_radius_m)
  movel([0.155811, -0.820667, -2.799119, -1.092603, 1.570796, 1.726607],accel_mss,speed_ms,0,blend_radius_m)
  movel([0.155954, -0.821400, -2.798989, -1.091999, 1.570796, 1.726751],accel_mss,speed_ms,0,blend_radius_m)
  movel([0.155514, -0.822266, -2.798836, -1.091287, 1.570796, 1.726310],accel_mss,speed_ms,0,blend_radius_m)
  movel([0.154880, -0.823093, -2.798689, -1.090607, 1.570796, 1.725676],accel_mss,speed_ms,0,blend_radius_m)
  movel([0.153372, -0.824368, -2.798461, -1.089559, 1.570796, 1.724168],accel_mss,speed_ms,0,blend_radius_m)
  movel([0.152148, -0.824931, -2.798361, -1.089097, 1.570796, 1.722944],accel_mss,speed_ms,0,blend_radius_m)
  movel([0.150940, -0.825247, -2.798304, -1.088838, 1.570796, 1.721736],accel_mss,speed_ms,0,blend_radius_m)
  movel([0.148664, -0.825648, -2.798232, -1.088509, 1.570796, 1.719461],accel_mss,speed_ms,0,blend_radius_m)
  movel([0.149487, -0.828629, -2.797695, -1.086065, 1.570796, 1.720283],accel_mss,speed_ms,0,blend_radius_m)
  movel([0.150580, -0.831339, -2.797203, -1.083847, 1.570796, 1.721377],accel_mss,speed_ms,0,blend_radius_m)
  movel([0.151941, -0.833766, -2.796759, -1.081864, 1.570796, 1.722738],accel_mss,speed_ms,0,blend_radius_m)
  movel([0.153547, -0.835914, -2.796363, -1.080112, 1.570796, 1.724344],accel_mss,speed_ms,0,blend_radius_m)
  movel([0.155518, -0.837569, -2.796056, -1.078764, 1.570796, 1.726315],accel_mss,speed_ms,0,blend_radius_m)
  movel([0.157892, -0.838681, -2.795849, -1.077859, 1.570796, 1.728688],accel_mss,speed_ms,0,blend_radius_m)
  movel([0.163164, -0.840120, -2.795580, -1.076689, 1.570796, 1.733961],accel_mss,speed_ms,0,blend_radius_m)
  movel([0.164477, -0.840859, -2.795442, -1.076088, 1.570796, 1.735273],accel_mss,speed_ms,0,blend_radius_m)
  movel([0.164731, -0.841607, -2.795301, -1.075481, 1.570796, 1.735527],accel_mss,speed_ms,0,blend_radius_m)
  movel([0.164486, -0.842690, -2.795097, -1.074602, 1.570796, 1.735282],accel_mss,speed_ms,0,blend_radius_m)
  movel([0.163859, -0.843737, -2.794899, -1.073752, 1.570796, 1.734656],accel_mss,speed_ms,0,blend_radius_m)
  movel([0.163012, -0.844665, -2.794724, -1.073000, 1.570796, 1.733808],accel_mss,speed_ms,0,blend_radius_m)
  movel([0.161071, -0.846127, -2.794446, -1.071816, 1.570796, 1.731867],accel_mss,speed_ms,0,blend_radius_m)
  movel([0.158538, -0.847537, -2.794177, -1.070675, 1.570796, 1.729334],accel_mss,speed_ms,0,blend_radius_m)
  movel([0.156117, -0.848591, -2.793975, -1.069824, 1.570796, 1.726913],accel_mss,speed_ms,0,blend_radius_m)
  movel([0.153793, -0.849345, -2.793830, -1.069214, 1.570796, 1.724589],accel_mss,speed_ms,0,blend_radius_m)
  movel([0.151559, -0.849834, -2.793736, -1.068819, 1.570796, 1.722355],accel_mss,speed_ms,0,blend_radius_m)
  movel([0.152827, -0.851880, -2.793340, -1.067168, 1.570796, 1.723624],accel_mss,speed_ms,0,blend_radius_m)
  movel([0.154404, -0.853545, -2.793017, -1.065827, 1.570796, 1.725200],accel_mss,speed_ms,0,blend_radius_m)
  movel([0.156283, -0.854784, -2.792775, -1.064830, 1.570796, 1.727080],accel_mss,speed_ms,0,blend_radius_m)
  movel([0.158458, -0.855563, -2.792623, -1.064203, 1.570796, 1.729255],accel_mss,speed_ms,0,blend_radius_m)
  movel([0.160934, -0.855833, -2.792570, -1.063986, 1.570796, 1.731730],accel_mss,speed_ms,0,blend_radius_m)
  movel([0.163710, -0.855556, -2.792624, -1.064208, 1.570796, 1.734507],accel_mss,speed_ms,0,blend_radius_m)
  movel([0.166787, -0.854683, -2.792795, -1.064911, 1.570796, 1.737583],accel_mss,speed_ms,0,blend_radius_m)
  movel([0.170171, -0.853170, -2.793090, -1.066129, 1.570796, 1.740967],accel_mss,speed_ms,0,blend_radius_m)
  speed_ms = 0.005
  movel([0.170171, -0.844130, -2.786876, -1.081383, 1.570796, 1.740967],accel_mss,speed_ms,0,blend_radius_m)
  speed_ms = 0.040
  movel([0.185325, -0.820896, -2.791208, -1.100285, 1.570796, 1.756121],accel_mss,speed_ms,0,blend_radius_m)
  speed_ms = 0.005
  movel([0.185325, -0.829723, -2.797497, -1.085169, 1.570796, 1.756121],accel_mss,speed_ms,0,blend_radius_m)
  speed_ms = 0.025
  movel([0.179130, -0.829569, -2.797525, -1.085295, 1.570796, 1.749926],accel_mss,speed_ms,0,blend_radius_m)
  movel([0.176504, -0.829194, -2.797593, -1.085602, 1.570796, 1.747300],accel_mss,speed_ms,0,blend_radius_m)
  movel([0.174175, -0.828518, -2.797716, -1.086156, 1.570796, 1.744971],accel_mss,speed_ms,0,blend_radius_m)
  movel([0.172123, -0.827457, -2.797907, -1.087025, 1.570796, 1.742919],accel_mss,speed_ms,0,blend_radius_m)
  movel([0.170335, -0.825936, -2.798181, -1.088273, 1.570796, 1.741131],accel_mss,speed_ms,0,blend_radius_m)
  movel([0.168788, -0.823879, -2.798549, -1.089961, 1.570796, 1.739584],accel_mss,speed_ms,0,blend_radius_m)
  movel([0.167475, -0.821202, -2.799024, -1.092162, 1.570796, 1.738271],accel_mss,speed_ms,0,blend_radius_m)
  movel([0.165467, -0.814874, -2.800134, -1.097381, 1.570796, 1.736263],accel_mss,speed_ms,0,blend_radius_m)
  movel([0.164156, -0.807856, -2.801339, -1.103194, 1.570796, 1.734952],accel_mss,speed_ms,0,blend_radius_m)
  movel([0.163481, -0.800234, -2.802619, -1.109536, 1.570796, 1.734277],accel_mss,speed_ms,0,blend_radius_m)
  movel([0.163370, -0.792111, -2.803951, -1.116327, 1.570796, 1.734166],accel_mss,speed_ms,0,blend_radius_m)
  movel([0.163693, -0.785112, -2.805071, -1.122206, 1.570796, 1.734489],accel_mss,speed_ms,0,blend_radius_m)
  movel([0.164351, -0.777836, -2.806210, -1.128343, 1.570796, 1.735147],accel_mss,speed_ms,0,blend_radius_m)
  movel([0.166427, -0.762599, -2.808510, -1.141280, 1.570796, 1.737223],accel_mss,speed_ms,0,blend_radius_m)
  movel([0.175526, -0.707594, -2.815904, -1.188890, 1.570796, 1.746322],accel_mss,speed_ms,0,blend_radius_m)
  movel([0.177448, -0.695750, -2.817317, -1.199321, 1.570796, 1.748244],accel_mss,speed_ms,0,blend_radius_m)
  movel([0.179180, -0.683923, -2.818668, -1.209798, 1.570796, 1.749976],accel_mss,speed_ms,0,blend_radius_m)
  movel([0.180554, -0.672288, -2.819938, -1.220162, 1.570796, 1.751350],accel_mss,speed_ms,0,blend_radius_m)
  movel([0.181390, -0.661014, -2.821115, -1.230260, 1.570796, 1.752186],accel_mss,speed_ms,0,blend_radius_m)
  movel([0.181508, -0.650289, -2.822186, -1.239913, 1.570796, 1.752305],accel_mss,speed_ms,0,blend_radius_m)
  movel([0.180716, -0.640314, -2.823140, -1.248935, 1.570796, 1.751512],accel_mss,speed_ms,0,blend_radius_m)
  movel([0.179492, -0.633612, -2.823759, -1.255018, 1.570796, 1.750288],accel_mss,speed_ms,0,blend_radius_m)
  movel([0.177674, -0.627254, -2.824329, -1.260806, 1.570796, 1.748470],accel_mss,speed_ms,0,blend_radius_m)
  movel([0.175212, -0.621422, -2.824838, -1.266129, 1.570796, 1.746008],accel_mss,speed_ms,0,blend_radius_m)
  movel([0.172054, -0.616298, -2.825274, -1.270816, 1.570796, 1.742851],accel_mss,speed_ms,0,blend_radius_m)
  movel([0.168163, -0.612056, -2.825628, -1.274705, 1.570796, 1.738959],accel_mss,speed_ms,0,blend_radius_m)
  movel([0.163499, -0.608866, -2.825889, -1.277634, 1.570796, 1.734295],accel_mss,speed_ms,0,blend_radius_m)
  movel([0.158021, -0.606916, -2.826047, -1.279426, 1.570796, 1.728817],accel_mss,speed_ms,0,blend_radius_m)
  movel([0.151716, -0.606363, -2.826091, -1.279935, 1.570796, 1.722513],accel_mss,speed_ms,0,blend_radius_m)
  movel([0.148431, -0.606690, -2.826065, -1.279634, 1.570796, 1.719227],accel_mss,speed_ms,0,blend_radius_m)
  movel([0.144882, -0.607482, -2.826001, -1.278906, 1.570796, 1.715678],accel_mss,speed_ms,0,blend_radius_m)
  movel([0.141095, -0.608759, -2.825898, -1.277732, 1.570796, 1.711892],accel_mss,speed_ms,0,blend_radius_m)
  movel([0.137112, -0.610533, -2.825753, -1.276103, 1.570796, 1.707908],accel_mss,speed_ms,0,blend_radius_m)
  movel([0.132975, -0.612800, -2.825566, -1.274023, 1.570796, 1.703772],accel_mss,speed_ms,0,blend_radius_m)
  movel([0.128708, -0.615588, -2.825334, -1.271467, 1.570796, 1.699505],accel_mss,speed_ms,0,blend_radius_m)
  movel([0.124362, -0.618885, -2.825055, -1.268448, 1.570796, 1.695159],accel_mss,speed_ms,0,blend_radius_m)
  movel([0.119974, -0.622707, -2.824727, -1.264955, 1.570796, 1.690770],accel_mss,speed_ms,0,blend_radius_m)
  speed_ms = 0.005
  movel([0.119974, -0.616589, -2.817929, -1.277871, 1.570796, 1.690770],accel_mss,speed_ms,0,blend_radius_m)
  speed_ms = 0.040
  movel([0.105668, -0.603740, -2.819005, -1.289644, 1.570796, 1.676464],accel_mss,speed_ms,0,blend_radius_m)
  speed_ms = 0.005
  movel([0.105668, -0.609641, -2.825826, -1.276922, 1.570796, 1.676464],accel_mss,speed_ms,0,blend_radius_m)
  speed_ms = 0.025
  movel([0.105208, -0.607230, -2.826021, -1.279138, 1.570796, 1.676004],accel_mss,speed_ms,0,blend_radius_m)
  movel([0.105101, -0.604506, -2.826240, -1.281644, 1.570796, 1.675897],accel_mss,speed_ms,0,blend_radius_m)
  movel([0.105749, -0.598322, -2.826724, -1.287343, 1.570796, 1.676545],accel_mss,speed_ms,0,blend_radius_m)
  movel([0.107230, -0.591444, -2.827246, -1.293698, 1.570796, 1.678026],accel_mss,speed_ms,0,blend_radius_m)
  movel([0.109136, -0.584270, -2.827772, -1.300347, 1.570796, 1.679932],accel_mss,speed_ms,0,blend_radius_m)
  speed_ms = 0.005
  movel([0.109136, -0.578803, -2.820912, -1.312675, 1.570796, 1.679932],accel_mss,speed_ms,0,blend_radius_m)
  speed_ms = 0.040
  movel([0.118580, -0.575376, -2.821155, -1.315858, 1.570796, 1.689376],accel_mss,speed_ms,0,blend_radius_m)
  speed_ms = 0.005
  movel([0.118580, -0.580783, -2.828020, -1.303586, 1.570796, 1.689376],accel_mss,speed_ms,0,blend_radius_m)
  speed_ms = 0.025
  movel([0.117402, -0.579337, -2.828122, -1.304930, 1.570796, 1.688198],accel_mss,speed_ms,0,blend_radius_m)
  movel([0.116582, -0.577565, -2.828246, -1.306579, 1.570796, 1.687379],accel_mss,speed_ms,0,blend_radius_m)
  movel([0.115918, -0.573127, -2.828550, -1.310712, 1.570796, 1.686715],accel_mss,speed_ms,0,blend_radius_m)
  movel([0.116427, -0.567666, -2.828915, -1.315809, 1.570796, 1.687223],accel_mss,speed_ms,0,blend_radius_m)
  movel([0.117944, -0.561360, -2.829322, -1.321707, 1.570796, 1.688741],accel_mss,speed_ms,0,blend_radius_m)
  movel([0.120304, -0.554407, -2.829754, -1.328228, 1.570796, 1.691100],accel_mss,speed_ms,0,blend_radius_m)
  movel([0.123332, -0.547011, -2.830194, -1.335184, 1.570796, 1.694129],accel_mss,speed_ms,0,blend_radius_m)
  movel([0.126853, -0.539377, -2.830628, -1.342384, 1.570796, 1.697649],accel_mss,speed_ms,0,blend_radius_m)
  movel([0.130680, -0.531724, -2.831042, -1.349622, 1.570796, 1.701476],accel_mss,speed_ms,0,blend_radius_m)
  speed_ms = 0.005
  movel([0.130680, -0.527205, -2.824113, -1.361071, 1.570796, 1.701476],accel_mss,speed_ms,0,blend_radius_m)
  speed_ms = 0.040
  movel([0.181260, -0.455421, -2.826978, -1.429990, 1.570796, 1.752057],accel_mss,speed_ms,0,blend_radius_m)
  speed_ms = 0.005
  movel([0.181260, -0.458521, -2.833970, -1.419898, 1.570796, 1.752057],accel_mss,speed_ms,0,blend_radius_m)
  speed_ms = 0.025
  movel([0.176078, -0.464566, -2.833797, -1.414025, 1.570796, 1.746874],accel_mss,speed_ms,0,blend_radius_m)
  movel([0.170926, -0.470930, -2.833603, -1.407856, 1.570796, 1.741722],accel_mss,speed_ms,0,blend_radius_m)
  movel([0.165890, -0.477510, -2.833387, -1.401492, 1.570796, 1.736686],accel_mss,speed_ms,0,blend_radius_m)
  movel([0.161028, -0.484229, -2.833152, -1.395008, 1.570796, 1.731824],accel_mss,speed_ms,0,blend_radius_m)
  movel([0.156423, -0.490997, -2.832899, -1.388494, 1.570796, 1.727219],accel_mss,speed_ms,0,blend_radius_m)
  movel([0.152136, -0.497723, -2.832632, -1.382034, 1.570796, 1.722932],accel_mss,speed_ms,0,blend_radius_m)
  movel([0.148234, -0.504335, -2.832354, -1.375700, 1.570796, 1.719030],accel_mss,speed_ms,0,blend_radius_m)
  movel([0.144778, -0.510756, -2.832070, -1.369563, 1.570796, 1.715575],accel_mss,speed_ms,0,blend_radius_m)
  movel([0.141828, -0.516899, -2.831785, -1.363705, 1.570796, 1.712624],accel_mss,speed_ms,0,blend_radius_m)
  movel([0.139435, -0.522705, -2.831504, -1.358181, 1.570796, 1.710232],accel_mss,speed_ms,0,blend_radius_m)
  movel([0.137657, -0.528098, -2.831231, -1.353060, 1.570796, 1.708453],accel_mss,speed_ms,0,blend_radius_m)
  movel([0.136544, -0.533010, -2.830974, -1.348405, 1.570796, 1.707340],accel_mss,speed_ms,0,blend_radius_m)
  movel([0.136155, -0.537371, -2.830739, -1.344279, 1.570796, 1.706952],accel_mss,speed_ms,0,blend_radius_m)
  movel([0.136543, -0.541117, -2.830531, -1.340741, 1.570796, 1.707339],accel_mss,speed_ms,0,blend_radius_m)
  movel([0.137752, -0.544189, -2.830357, -1.337843, 1.570796, 1.708548],accel_mss,speed_ms,0,blend_radius_m)
  movel([0.139843, -0.546520, -2.830223, -1.335646, 1.570796, 1.710639],accel_mss,speed_ms,0,blend_radius_m)
  speed_ms = 0.005
  movel([0.139843, -0.541727, -2.823311, -1.347350, 1.570796, 1.710639],accel_mss,speed_ms,0,blend_radius_m)
  speed_ms = 0.040
  movel([0.162855, -0.515901, -2.824685, -1.371803, 1.570796, 1.733652],accel_mss,speed_ms,0,blend_radius_m)
  speed_ms = 0.005
  movel([0.162855, -0.520204, -2.831626, -1.360559, 1.570796, 1.733652],accel_mss,speed_ms,0,blend_radius_m)
  speed_ms = 0.025
  movel([0.162384, -0.517247, -2.831769, -1.363373, 1.570796, 1.733180],accel_mss,speed_ms,0,blend_radius_m)
  movel([0.162288, -0.513923, -2.831925, -1.366541, 1.570796, 1.733084],accel_mss,speed_ms,0,blend_radius_m)
  movel([0.162565, -0.510268, -2.832093, -1.370028, 1.570796, 1.733362],accel_mss,speed_ms,0,blend_radius_m)
  movel([0.163216, -0.506303, -2.832269, -1.373817, 1.570796, 1.734012],accel_mss,speed_ms,0,blend_radius_m)
  movel([0.164233, -0.502063, -2.832452, -1.377874, 1.570796, 1.735029],accel_mss,speed_ms,0,blend_radius_m)
  movel([0.165623, -0.497570, -2.832638, -1.382181, 1.570796, 1.736419],accel_mss,speed_ms,0,blend_radius_m)
  movel([0.167387, -0.492843, -2.832827, -1.386719, 1.570796, 1.738183],accel_mss,speed_ms,0,blend_radius_m)
  movel([0.169516, -0.487927, -2.833015, -1.391447, 1.570796, 1.740313],accel_mss,speed_ms,0,blend_radius_m)
  movel([0.172012, -0.482842, -2.833201, -1.396346, 1.570796, 1.742809],accel_mss,speed_ms,0,blend_radius_m)
  movel([0.174881, -0.477611, -2.833384, -1.401395, 1.570796, 1.745678],accel_mss,speed_ms,0,blend_radius_m)
  movel([0.178106, -0.472287, -2.833559, -1.406543, 1.570796, 1.748902],accel_mss,speed_ms,0,blend_radius_m)
  movel([0.181701, -0.466876, -2.833728, -1.411785, 1.570796, 1.752497],accel_mss,speed_ms,0,blend_radius_m)
  movel([0.185655, -0.461422, -2.833888, -1.417079, 1.570796, 1.756451],accel_mss,speed_ms,0,blend_radius_m)
  movel([0.189965, -0.455956, -2.834039, -1.422394, 1.570796, 1.760761],accel_mss,speed_ms,0,blend_radius_m)
  movel([0.194624, -0.450521, -2.834179, -1.427690, 1.570796, 1.765421],accel_mss,speed_ms,0,blend_radius_m)
  movel([0.199621, -0.445150, -2.834307, -1.432932, 1.570796, 1.770417],accel_mss,speed_ms,0,blend_radius_m)
  movel([0.204634, -0.440209, -2.834417, -1.437763, 1.570796, 1.775430],accel_mss,speed_ms,0,blend_radius_m)
  movel([0.209620, -0.435725, -2.834509, -1.442155, 1.570796, 1.780416],accel_mss,speed_ms,0,blend_radius_m)
  movel([0.214539, -0.431701, -2.834586, -1.446102, 1.570796, 1.785336],accel_mss,speed_ms,0,blend_radius_m)
  movel([0.219373, -0.428139, -2.834650, -1.449600, 1.570796, 1.790170],accel_mss,speed_ms,0,blend_radius_m)
  movel([0.224084, -0.425042, -2.834702, -1.452645, 1.570796, 1.794880],accel_mss,speed_ms,0,blend_radius_m)
  movel([0.228628, -0.422427, -2.834744, -1.455219, 1.570796, 1.799425],accel_mss,speed_ms,0,blend_radius_m)
  movel([0.232995, -0.420270, -2.834776, -1.457343, 1.570796, 1.803792],accel_mss,speed_ms,0,blend_radius_m)
  movel([0.237129, -0.418598, -2.834801, -1.458991, 1.570796, 1.807925],accel_mss,speed_ms,0,blend_radius_m)
  movel([0.241016, -0.417398, -2.834817, -1.460174, 1.570796, 1.811812],accel_mss,speed_ms,0,blend_radius_m)
  movel([0.247935, -0.416393, -2.834831, -1.461165, 1.570796, 1.818732],accel_mss,speed_ms,0,blend_radius_m)
  movel([0.250900, -0.416592, -2.834828, -1.460968, 1.570796, 1.821697],accel_mss,speed_ms,0,blend_radius_m)
  movel([0.255753, -0.418336, -2.834804, -1.459249, 1.570796, 1.826549],accel_mss,speed_ms,0,blend_radius_m)
  movel([0.257590, -0.419864, -2.834782, -1.457743, 1.570796, 1.828387],accel_mss,speed_ms,0,blend_radius_m)
  movel([0.259001, -0.421823, -2.834753, -1.455813, 1.570796, 1.829798],accel_mss,speed_ms,0,blend_radius_m)
  speed_ms = 0.005
  movel([0.259001, -0.419469, -2.827745, -1.465175, 1.570796, 1.829798],accel_mss,speed_ms,0,blend_radius_m)
  speed_ms = 0.040
  movel([0.274724, -0.432636, -2.827515, -1.452238, 1.570796, 1.845520],accel_mss,speed_ms,0,blend_radius_m)
  speed_ms = 0.005
  movel([0.274724, -0.435265, -2.834518, -1.442606, 1.570796, 1.845520],accel_mss,speed_ms,0,blend_radius_m)
  speed_ms = 0.025
  movel([0.272812, -0.432026, -2.834580, -1.445783, 1.570796, 1.843609],accel_mss,speed_ms,0,blend_radius_m)
  movel([0.269936, -0.429968, -2.834618, -1.447803, 1.570796, 1.840732],accel_mss,speed_ms,0,blend_radius_m)
  movel([0.266170, -0.429088, -2.834633, -1.448667, 1.570796, 1.836967],accel_mss,speed_ms,0,blend_radius_m)
  movel([0.261578, -0.429385, -2.834628, -1.448376, 1.570796, 1.832374],accel_mss,speed_ms,0,blend_radius_m)
  movel([0.256264, -0.430831, -2.834602, -1.446956, 1.570796, 1.827060],accel_mss,speed_ms,0,blend_radius_m)
  movel([0.250302, -0.433418, -2.834554, -1.444418, 1.570796, 1.821099],accel_mss,speed_ms,0,blend_radius_m)
  movel([0.243802, -0.437109, -2.834481, -1.440799, 1.570796, 1.814599],accel_mss,speed_ms,0,blend_radius_m)
  movel([0.236850, -0.441880, -2.834380, -1.436129, 1.570796, 1.807647],accel_mss,speed_ms,0,blend_radius_m)
  movel([0.229570, -0.447678, -2.834248, -1.430464, 1.570796, 1.800366],accel_mss,speed_ms,0,blend_radius_m)
  movel([0.222137, -0.454386, -2.834080, -1.423923, 1.570796, 1.792933],accel_mss,speed_ms,0,blend_radius_m)
  movel([0.214847, -0.461760, -2.833879, -1.416750, 1.570796, 1.785644],accel_mss,speed_ms,0,blend_radius_m)
  movel([0.208004, -0.469563, -2.833646, -1.409180, 1.570796, 1.778801],accel_mss,speed_ms,0,blend_radius_m)
  movel([0.201871, -0.477580, -2.833385, -1.401424, 1.570796, 1.772667],accel_mss,speed_ms,0,blend_radius_m)
  movel([0.199162, -0.481595, -2.833246, -1.397548, 1.570796, 1.769958],accel_mss,speed_ms,0,blend_radius_m)
  movel([0.196726, -0.485580, -2.833102, -1.393707, 1.570796, 1.767523],accel_mss,speed_ms,0,blend_radius_m)
  movel([0.194595, -0.489515, -2.832955, -1.389919, 1.570796, 1.765391],accel_mss,speed_ms,0,blend_radius_m)
  movel([0.192805, -0.493375, -2.832806, -1.386207, 1.570796, 1.763601],accel_mss,speed_ms,0,blend_radius_m)
  movel([0.191376, -0.497135, -2.832656, -1.382598, 1.570796, 1.762173],accel_mss,speed_ms,0,blend_radius_m)
  movel([0.190353, -0.500760, -2.832506, -1.379122, 1.570796, 1.761149],accel_mss,speed_ms,0,blend_radius_m)
  speed_ms = 0.005
  movel([0.190353, -0.496829, -2.825547, -1.390014, 1.570796, 1.761149],accel_mss,speed_ms,0,blend_radius_m)
  speed_ms = 0.040
  movel([0.225557, -0.485564, -2.825995, -1.400830, 1.570796, 1.796354],accel_mss,speed_ms,0,blend_radius_m)
  speed_ms = 0.005
  movel([0.225557, -0.489272, -2.832965, -1.390152, 1.570796, 1.796354],accel_mss,speed_ms,0,blend_radius_m)
  speed_ms = 0.025
  movel([0.230532, -0.483646, -2.833173, -1.395570, 1.570796, 1.801329],accel_mss,speed_ms,0,blend_radius_m)
  movel([0.235675, -0.478496, -2.833353, -1.400539, 1.570796, 1.806472],accel_mss,speed_ms,0,blend_radius_m)
  movel([0.240904, -0.473851, -2.833509, -1.405029, 1.570796, 1.811700],accel_mss,speed_ms,0,blend_radius_m)
  movel([0.246113, -0.469761, -2.833639, -1.408988, 1.570796, 1.816909],accel_mss,speed_ms,0,blend_radius_m)
  movel([0.251210, -0.466259, -2.833747, -1.412383, 1.570796, 1.822007],accel_mss,speed_ms,0,blend_radius_m)
  movel([0.256093, -0.463379, -2.833832, -1.415178, 1.570796, 1.826889],accel_mss,speed_ms,0,blend_radius_m)
  movel([0.260676, -0.461152, -2.833896, -1.417340, 1.570796, 1.831472],accel_mss,speed_ms,0,blend_radius_m)
  movel([0.264851, -0.459614, -2.833939, -1.418836, 1.570796, 1.835647],accel_mss,speed_ms,0,blend_radius_m)
  movel([0.269216, -0.458845, -2.833961, -1.419583, 1.570796, 1.840012],accel_mss,speed_ms,0,blend_radius_m)
  movel([0.272323, -0.459454, -2.833944, -1.418991, 1.570796, 1.843120],accel_mss,speed_ms,0,blend_radius_m)
  movel([0.274310, -0.461289, -2.833892, -1.417208, 1.570796, 1.845106],accel_mss,speed_ms,0,blend_radius_m)
  movel([0.275291, -0.464214, -2.833808, -1.414367, 1.570796, 1.846087],accel_mss,speed_ms,0,blend_radius_m)
  movel([0.275404, -0.468063, -2.833692, -1.410634, 1.570796, 1.846201],accel_mss,speed_ms,0,blend_radius_m)
  movel([0.274782, -0.472696, -2.833546, -1.406146, 1.570796, 1.845579],accel_mss,speed_ms,0,blend_radius_m)
  movel([0.273555, -0.477960, -2.833372, -1.401057, 1.570796, 1.844351],accel_mss,speed_ms,0,blend_radius_m)
  movel([0.271863, -0.483700, -2.833171, -1.395518, 1.570796, 1.842660],accel_mss,speed_ms,0,blend_radius_m)
  speed_ms = 0.005
  movel([0.271863, -0.480100, -2.826197, -1.406092, 1.570796, 1.842660],accel_mss,speed_ms,0,blend_radius_m)
  speed_ms = 0.040
  movel([0.237934, -0.500739, -2.825380, -1.386269, 1.570796, 1.808730],accel_mss,speed_ms,0,blend_radius_m)
  speed_ms = 0.005
  movel([0.237934, -0.504748, -2.832337, -1.375305, 1.570796, 1.808730],accel_mss,speed_ms,0,blend_radius_m)
  speed_ms = 0.025
  movel([0.242451, -0.502306, -2.832441, -1.377641, 1.570796, 1.813247],accel_mss,speed_ms,0,blend_radius_m)
  movel([0.246530, -0.500594, -2.832513, -1.379282, 1.570796, 1.817326],accel_mss,speed_ms,0,blend_radius_m)
  movel([0.250167, -0.499593, -2.832555, -1.380241, 1.570796, 1.820964],accel_mss,speed_ms,0,blend_radius_m)
  movel([0.253371, -0.499255, -2.832569, -1.380565, 1.570796, 1.824168],accel_mss,speed_ms,0,blend_radius_m)
  movel([0.256145, -0.499552, -2.832557, -1.380280, 1.570796, 1.826941],accel_mss,speed_ms,0,blend_radius_m)
  movel([0.258492, -0.500442, -2.832520, -1.379428, 1.570796, 1.829288],accel_mss,speed_ms,0,blend_radius_m)
  movel([0.260428, -0.501883, -2.832459, -1.378047, 1.570796, 1.831224],accel_mss,speed_ms,0,blend_radius_m)
  movel([0.261949, -0.503847, -2.832375, -1.376166, 1.570796, 1.832745],accel_mss,speed_ms,0,blend_radius_m)
  movel([0.263082, -0.506281, -2.832270, -1.373838, 1.570796, 1.833878],accel_mss,speed_ms,0,blend_radius_m)
  movel([0.263834, -0.509144, -2.832143, -1.371102, 1.570796, 1.834630],accel_mss,speed_ms,0,blend_radius_m)
  movel([0.264212, -0.512402, -2.831995, -1.367992, 1.570796, 1.835008],accel_mss,speed_ms,0,blend_radius_m)
  movel([0.264237, -0.516002, -2.831828, -1.364559, 1.570796, 1.835033],accel_mss,speed_ms,0,blend_radius_m)
  movel([0.263917, -0.519912, -2.831641, -1.360836, 1.570796, 1.834713],accel_mss,speed_ms,0,blend_radius_m)
  movel([0.262305, -0.528475, -2.831212, -1.352702, 1.570796, 1.833101],accel_mss,speed_ms,0,blend_radius_m)
  movel([0.261033, -0.533057, -2.830972, -1.348360, 1.570796, 1.831830],accel_mss,speed_ms,0,blend_radius_m)
  movel([0.260911, -0.531907, -2.831033, -1.349449, 1.570796, 1.831708],accel_mss,speed_ms,0,blend_radius_m)
  speed_ms = 0.005
  movel([0.260911, -0.527384, -2.824104, -1.360900, 1.570796, 1.831708],accel_mss,speed_ms,0,blend_radius_m)
  speed_ms = 0.040
  movel([0.286425, -0.525905, -2.824182, -1.362302, 1.570796, 1.857221],accel_mss,speed_ms,0,blend_radius_m)
  speed_ms = 0.005
  movel([0.286425, -0.530400, -2.831112, -1.350877, 1.570796, 1.857221],accel_mss,speed_ms,0,blend_radius_m)
  speed_ms = 0.025
  movel([0.281721, -0.537880, -2.830711, -1.343798, 1.570796, 1.852517],accel_mss,speed_ms,0,blend_radius_m)
  movel([0.277579, -0.545251, -2.830296, -1.336842, 1.570796, 1.848375],accel_mss,speed_ms,0,blend_radius_m)
  movel([0.273882, -0.552492, -2.829870, -1.330027, 1.570796, 1.844679],accel_mss,speed_ms,0,blend_radius_m)
  movel([0.270506, -0.559590, -2.829433, -1.323366, 1.570796, 1.841302],accel_mss,speed_ms,0,blend_radius_m)
  movel([0.267119, -0.567242, -2.828942, -1.316205, 1.570796, 1.837915],accel_mss,speed_ms,0,blend_radius_m)
  movel([0.265729, -0.570898, -2.828700, -1.312791, 1.570796, 1.836525],accel_mss,speed_ms,0,blend_radius_m)
  movel([0.264664, -0.574360, -2.828466, -1.309563, 1.570796, 1.835460],accel_mss,speed_ms,0,blend_radius_m)
  movel([0.264005, -0.577559, -2.828246, -1.306584, 1.570796, 1.834801],accel_mss,speed_ms,0,blend_radius_m)
  movel([0.263849, -0.580357, -2.828051, -1.303981, 1.570796, 1.834645],accel_mss,speed_ms,0,blend_radius_m)
  movel([0.264284, -0.582577, -2.827893, -1.301919, 1.570796, 1.835080],accel_mss,speed_ms,0,blend_radius_m)
  movel([0.265378, -0.584075, -2.827786, -1.300528, 1.570796, 1.836174],accel_mss,speed_ms,0,blend_radius_m)
  movel([0.268144, -0.585109, -2.827712, -1.299569, 1.570796, 1.838940],accel_mss,speed_ms,0,blend_radius_m)
  movel([0.269503, -0.585645, -2.827673, -1.299071, 1.570796, 1.840299],accel_mss,speed_ms,0,blend_radius_m)
  movel([0.270510, -0.586622, -2.827602, -1.298165, 1.570796, 1.841306],accel_mss,speed_ms,0,blend_radius_m)
  movel([0.270926, -0.588607, -2.827457, -1.296326, 1.570796, 1.841723],accel_mss,speed_ms,0,blend_radius_m)
  movel([0.270622, -0.591459, -2.827245, -1.293684, 1.570796, 1.841419],accel_mss,speed_ms,0,blend_radius_m)
  movel([0.269763, -0.594946, -2.826983, -1.290460, 1.570796, 1.840560],accel_mss,speed_ms,0,blend_radius_m)
  movel([0.268504, -0.598829, -2.826685, -1.286875, 1.570796, 1.839300],accel_mss,speed_ms,0,blend_radius_m)
  movel([0.265395, -0.606888, -2.826049, -1.279452, 1.570796, 1.836191],accel_mss,speed_ms,0,blend_radius_m)
  movel([0.255783, -0.629500, -2.824129, -1.258760, 1.570796, 1.826579],accel_mss,speed_ms,0,blend_radius_m)
  movel([0.249309, -0.644871, -2.822710, -1.244809, 1.570796, 1.820106],accel_mss,speed_ms,0,blend_radius_m)
  movel([0.247618, -0.649444, -2.822269, -1.240676, 1.570796, 1.818415],accel_mss,speed_ms,0,blend_radius_m)
  movel([0.246095, -0.654195, -2.821802, -1.236392, 1.570796, 1.816891],accel_mss,speed_ms,0,blend_radius_m)
  movel([0.243703, -0.663807, -2.820829, -1.227753, 1.570796, 1.814500],accel_mss,speed_ms,0,blend_radius_m)
  movel([0.242917, -0.668461, -2.820344, -1.223584, 1.570796, 1.813713],accel_mss,speed_ms,0,blend_radius_m)
  movel([0.242456, -0.672873, -2.819876, -1.219640, 1.570796, 1.813252],accel_mss,speed_ms,0,blend_radius_m)
  movel([0.242353, -0.676948, -2.819437, -1.216005, 1.570796, 1.813149],accel_mss,speed_ms,0,blend_radius_m)
  movel([0.242645, -0.680589, -2.819038, -1.212762, 1.570796, 1.813442],accel_mss,speed_ms,0,blend_radius_m)
  movel([0.243374, -0.683688, -2.818694, -1.210007, 1.570796, 1.814170],accel_mss,speed_ms,0,blend_radius_m)
  movel([0.244568, -0.686166, -2.818416, -1.207806, 1.570796, 1.815364],accel_mss,speed_ms,0,blend_radius_m)
  movel([0.246276, -0.687910, -2.818219, -1.206259, 1.570796, 1.817072],accel_mss,speed_ms,0,blend_radius_m)
  movel([0.248533, -0.688829, -2.818115, -1.205445, 1.570796, 1.819329],accel_mss,speed_ms,0,blend_radius_m)
  movel([0.251378, -0.688824, -2.818116, -1.205449, 1.570796, 1.822174],accel_mss,speed_ms,0,blend_radius_m)
  movel([0.254864, -0.687787, -2.818233, -1.206369, 1.570796, 1.825661],accel_mss,speed_ms,0,blend_radius_m)
  movel([0.259038, -0.685617, -2.818478, -1.208294, 1.570796, 1.829835],accel_mss,speed_ms,0,blend_radius_m)
  movel([0.263958, -0.682198, -2.818860, -1.211331, 1.570796, 1.834754],accel_mss,speed_ms,0,blend_radius_m)
  movel([0.267886, -0.678956, -2.819217, -1.214215, 1.570796, 1.838682],accel_mss,speed_ms,0,blend_radius_m)
  movel([0.271783, -0.675350, -2.819610, -1.217429, 1.570796, 1.842579],accel_mss,speed_ms,0,blend_radius_m)
  movel([0.275661, -0.671427, -2.820030, -1.220931, 1.570796, 1.846457],accel_mss,speed_ms,0,blend_radius_m)
  movel([0.279521, -0.667250, -2.820471, -1.224668, 1.570796, 1.850318],accel_mss,speed_ms,0,blend_radius_m)
  movel([0.287206, -0.658376, -2.821383, -1.232630, 1.570796, 1.858002],accel_mss,speed_ms,0,blend_radius_m)
  movel([0.294865, -0.649219, -2.822291, -1.240879, 1.570796, 1.865661],accel_mss,speed_ms,0,blend_radius_m)
  movel([0.302757, -0.640072, -2.823163, -1.249154, 1.570796, 1.873553],accel_mss,speed_ms,0,blend_radius_m)
  movel([0.306845, -0.635614, -2.823576, -1.253199, 1.570796, 1.877642],accel_mss,speed_ms,0,blend_radius_m)
  movel([0.310988, -0.631365, -2.823962, -1.257061, 1.570796, 1.881784],accel_mss,speed_ms,0,blend_radius_m)
  movel([0.315153, -0.627410, -2.824315, -1.260664, 1.570796, 1.885950],accel_mss,speed_ms,0,blend_radius_m)
  movel([0.319307, -0.623855, -2.824627, -1.263906, 1.570796, 1.890104],accel_mss,speed_ms,0,blend_radius_m)
  movel([0.323408, -0.620799, -2.824892, -1.266698, 1.570796, 1.894204],accel_mss,speed_ms,0,blend_radius_m)
  movel([0.327424, -0.618343, -2.825101, -1.268944, 1.570796, 1.898220],accel_mss,speed_ms,0,blend_radius_m)
  movel([0.335704, -0.614576, -2.825419, -1.272394, 1.570796, 1.906501],accel_mss,speed_ms,0,blend_radius_m)
  movel([0.338553, -0.613069, -2.825544, -1.273776, 1.570796, 1.909349],accel_mss,speed_ms,0,blend_radius_m)
  movel([0.341622, -0.610968, -2.825717, -1.275703, 1.570796, 1.912418],accel_mss,speed_ms,0,blend_radius_m)
  movel([0.344775, -0.608229, -2.825941, -1.278219, 1.570796, 1.915572],accel_mss,speed_ms,0,blend_radius_m)
  movel([0.347727, -0.604986, -2.826201, -1.281202, 1.570796, 1.918524],accel_mss,speed_ms,0,blend_radius_m)
  movel([0.349043, -0.603209, -2.826342, -1.282837, 1.570796, 1.919839],accel_mss,speed_ms,0,blend_radius_m)
  movel([0.350203, -0.601354, -2.826489, -1.284546, 1.570796, 1.920999],accel_mss,speed_ms,0,blend_radius_m)
  speed_ms = 0.005
  movel([0.350203, -0.595593, -2.819654, -1.297141, 1.570796, 1.920999],accel_mss,speed_ms,0,blend_radius_m)
  speed_ms = 0.040
  movel([0.368105, -0.561778, -2.822077, -1.328534, 1.570796, 1.938901],accel_mss,speed_ms,0,blend_radius_m)
  speed_ms = 0.005
  movel([0.368105, -0.566940, -2.828962, -1.316486, 1.570796, 1.938901],accel_mss,speed_ms,0,blend_radius_m)
  speed_ms = 0.025
  movel([0.368968, -0.567013, -2.828957, -1.316418, 1.570796, 1.939765],accel_mss,speed_ms,0,blend_radius_m)
  movel([0.368864, -0.568264, -2.828875, -1.315250, 1.570796, 1.939660],accel_mss,speed_ms,0,blend_radius_m)
  movel([0.368010, -0.570104, -2.828753, -1.313532, 1.570796, 1.938806],accel_mss,speed_ms,0,blend_radius_m)
  movel([0.366650, -0.571947, -2.828630, -1.311812, 1.570796, 1.937447],accel_mss,speed_ms,0,blend_radius_m)
  movel([0.365112, -0.573388, -2.828532, -1.310469, 1.570796, 1.935908],accel_mss,speed_ms,0,blend_radius_m)
  movel([0.363581, -0.574513, -2.828456, -1.309420, 1.570796, 1.934377],accel_mss,speed_ms,0,blend_radius_m)
  movel([0.360546, -0.576432, -2.828324, -1.307633, 1.570796, 1.931342],accel_mss,speed_ms,0,blend_radius_m)
  movel([0.358317, -0.578078, -2.828210, -1.306101, 1.570796, 1.929113],accel_mss,speed_ms,0,blend_radius_m)
  movel([0.356086, -0.580022, -2.828074, -1.304293, 1.570796, 1.926882],accel_mss,speed_ms,0,blend_radius_m)
  movel([0.351647, -0.584587, -2.827749, -1.300053, 1.570796, 1.922443],accel_mss,speed_ms,0,blend_radius_m)
  movel([0.347317, -0.589717, -2.827375, -1.295297, 1.570796, 1.918113],accel_mss,speed_ms,0,blend_radius_m)
  movel([0.343182, -0.594983, -2.826980, -1.290426, 1.570796, 1.913979],accel_mss,speed_ms,0,blend_radius_m)
  movel([0.342235, -0.596290, -2.826881, -1.289219, 1.570796, 1.913032],accel_mss,speed_ms,0,blend_radius_m)
  movel([0.341615, -0.597527, -2.826786, -1.288076, 1.570796, 1.912411],accel_mss,speed_ms,0,blend_radius_m)
  movel([0.341723, -0.598419, -2.826717, -1.287253, 1.570796, 1.912520],accel_mss,speed_ms,0,blend_radius_m)
  movel([0.342462, -0.598661, -2.826698, -1.287030, 1.570796, 1.913258],accel_mss,speed_ms,0,blend_radius_m)
  movel([0.344503, -0.598547, -2.826707, -1.287135, 1.570796, 1.915299],accel_mss,speed_ms,0,blend_radius_m)
  movel([0.346807, -0.597940, -2.826754, -1.287695, 1.570796, 1.917604],accel_mss,speed_ms,0,blend_radius_m)
  movel([0.349334, -0.596873, -2.826836, -1.288680, 1.570796, 1.920130],accel_mss,speed_ms,0,blend_radius_m)
  movel([0.352037, -0.595364, -2.826951, -1.290074, 1.570796, 1.922833],accel_mss,speed_ms,0,blend_radius_m)
  movel([0.354856, -0.593461, -2.827095, -1.291833, 1.570796, 1.925652],accel_mss,speed_ms,0,blend_radius_m)
  movel([0.357752, -0.591175, -2.827267, -1.293948, 1.570796, 1.928549],accel_mss,speed_ms,0,blend_radius_m)
  movel([0.360668, -0.588549, -2.827461, -1.296379, 1.570796, 1.931464],accel_mss,speed_ms,0,blend_radius_m)
  movel([0.363561, -0.585598, -2.827676, -1.299115, 1.570796, 1.934358],accel_mss,speed_ms,0,blend_radius_m)
  movel([0.362934, -0.587425, -2.827543, -1.297421, 1.570796, 1.933731],accel_mss,speed_ms,0,blend_radius_m)
  movel([0.363038, -0.588714, -2.827449, -1.296226, 1.570796, 1.933835],accel_mss,speed_ms,0,blend_radius_m)
  movel([0.363749, -0.589393, -2.827399, -1.295597, 1.570796, 1.934545],accel_mss,speed_ms,0,blend_radius_m)
  movel([0.364933, -0.589393, -2.827399, -1.295597, 1.570796, 1.935729],accel_mss,speed_ms,0,blend_radius_m)
  movel([0.366423, -0.588768, -2.827445, -1.296176, 1.570796, 1.937220],accel_mss,speed_ms,0,blend_radius_m)
  movel([0.368082, -0.587710, -2.827522, -1.297157, 1.570796, 1.938878],accel_mss,speed_ms,0,blend_radius_m)
  movel([0.371589, -0.584790, -2.827735, -1.299865, 1.570796, 1.942385],accel_mss,speed_ms,0,blend_radius_m)
  movel([0.376077, -0.580358, -2.828050, -1.303980, 1.570796, 1.946874],accel_mss,speed_ms,0,blend_radius_m)
  movel([0.380438, -0.575425, -2.828393, -1.308571, 1.570796, 1.951234],accel_mss,speed_ms,0,blend_radius_m)
  movel([0.384550, -0.570139, -2.828751, -1.313499, 1.570796, 1.955347],accel_mss,speed_ms,0,blend_radius_m)
  movel([0.388290, -0.564643, -2.829112, -1.318634, 1.570796, 1.959086],accel_mss,speed_ms,0,blend_radius_m)
  movel([0.389384, -0.562776, -2.829232, -1.320381, 1.570796, 1.960180],accel_mss,speed_ms,0,blend_radius_m)
  movel([0.389964, -0.561155, -2.829335, -1.321899, 1.570796, 1.960761],accel_mss,speed_ms,0,blend_radius_m)
  movel([0.389788, -0.560315, -2.829388, -1.322686, 1.570796, 1.960584],accel_mss,speed_ms,0,blend_radius_m)
  movel([0.389203, -0.559913, -2.829413, -1.323063, 1.570796, 1.959999],accel_mss,speed_ms,0,blend_radius_m)
  movel([0.386676, -0.559370, -2.829447, -1.323571, 1.570796, 1.957472],accel_mss,speed_ms,0,blend_radius_m)
  movel([0.381451, -0.559187, -2.829459, -1.323743, 1.570796, 1.952247],accel_mss,speed_ms,0,blend_radius_m)
  movel([0.379326, -0.558064, -2.829529, -1.324796, 1.570796, 1.950122],accel_mss,speed_ms,0,blend_radius_m)
  movel([0.384469, -0.551946, -2.829903, -1.330540, 1.570796, 1.955266],accel_mss,speed_ms,0,blend_radius_m)
  movel([0.387180, -0.549202, -2.830066, -1.333121, 1.570796, 1.957976],accel_mss,speed_ms,0,blend_radius_m)
  movel([0.389910, -0.546850, -2.830204, -1.335335, 1.570796, 1.960706],accel_mss,speed_ms,0,blend_radius_m)
  movel([0.391735, -0.545577, -2.830277, -1.336534, 1.570796, 1.962531],accel_mss,speed_ms,0,blend_radius_m)
  movel([0.393582, -0.544545, -2.830337, -1.337507, 1.570796, 1.964378],accel_mss,speed_ms,0,blend_radius_m)
  movel([0.396744, -0.543462, -2.830399, -1.338528, 1.570796, 1.967540],accel_mss,speed_ms,0,blend_radius_m)
  movel([0.398201, -0.543893, -2.830374, -1.338122, 1.570796, 1.968997],accel_mss,speed_ms,0,blend_radius_m)
  movel([0.398494, -0.544631, -2.830332, -1.337426, 1.570796, 1.969291],accel_mss,speed_ms,0,blend_radius_m)
  movel([0.398393, -0.545741, -2.830268, -1.336380, 1.570796, 1.969189],accel_mss,speed_ms,0,blend_radius_m)
  movel([0.397663, -0.547579, -2.830161, -1.334649, 1.570796, 1.968460],accel_mss,speed_ms,0,blend_radius_m)
  movel([0.396447, -0.549587, -2.830043, -1.332759, 1.570796, 1.967243],accel_mss,speed_ms,0,blend_radius_m)
  movel([0.393297, -0.553609, -2.829802, -1.328978, 1.570796, 1.964093],accel_mss,speed_ms,0,blend_radius_m)
  speed_ms = 0.005
  movel([0.393297, -0.548686, -2.822900, -1.340803, 1.570796, 1.964093],accel_mss,speed_ms,0,blend_radius_m)
  speed_ms = 0.040
  movel([0.440057, -0.419703, -2.827741, -1.464944, 1.570796, 2.010854],accel_mss,speed_ms,0,blend_radius_m)
  speed_ms = 0.005
  movel([0.440057, -0.422062, -2.834749, -1.455578, 1.570796, 2.010854],accel_mss,speed_ms,0,blend_radius_m)
  speed_ms = 0.025
  movel([0.442441, -0.419837, -2.834783, -1.457770, 1.570796, 2.013238],accel_mss,speed_ms,0,blend_radius_m)
  movel([0.444761, -0.417990, -2.834809, -1.459590, 1.570796, 2.015558],accel_mss,speed_ms,0,blend_radius_m)
  movel([0.446970, -0.416528, -2.834829, -1.461031, 1.570796, 2.017767],accel_mss,speed_ms,0,blend_radius_m)
  movel([0.450910, -0.414773, -2.834852, -1.462764, 1.570796, 2.021706],accel_mss,speed_ms,0,blend_radius_m)
  movel([0.452557, -0.414482, -2.834856, -1.463050, 1.570796, 2.023353],accel_mss,speed_ms,0,blend_radius_m)
  movel([0.455003, -0.415089, -2.834848, -1.462452, 1.570796, 2.025800],accel_mss,speed_ms,0,blend_radius_m)
  movel([0.456272, -0.417086, -2.834822, -1.460481, 1.570796, 2.027069],accel_mss,speed_ms,0,blend_radius_m)
  movel([0.456587, -0.420094, -2.834779, -1.457517, 1.570796, 2.027383],accel_mss,speed_ms,0,blend_radius_m)
  movel([0.456142, -0.423840, -2.834722, -1.453828, 1.570796, 2.026938],accel_mss,speed_ms,0,blend_radius_m)
  movel([0.455131, -0.428055, -2.834652, -1.449683, 1.570796, 2.025928],accel_mss,speed_ms,0,blend_radius_m)
  movel([0.452847, -0.434973, -2.834524, -1.442892, 1.570796, 2.023643],accel_mss,speed_ms,0,blend_radius_m)
  movel([0.449787, -0.442383, -2.834369, -1.435637, 1.570796, 2.020584],accel_mss,speed_ms,0,blend_radius_m)
  movel([0.446023, -0.450150, -2.834188, -1.428051, 1.570796, 2.016820],accel_mss,speed_ms,0,blend_radius_m)
  movel([0.437383, -0.465709, -2.833763, -1.412917, 1.570796, 2.008179],accel_mss,speed_ms,0,blend_radius_m)
  movel([0.435923, -0.469076, -2.833661, -1.409652, 1.570796, 2.006720],accel_mss,speed_ms,0,blend_radius_m)
  movel([0.435426, -0.471753, -2.833577, -1.407060, 1.570796, 2.006222],accel_mss,speed_ms,0,blend_radius_m)
  movel([0.435982, -0.473233, -2.833529, -1.405627, 1.570796, 2.006778],accel_mss,speed_ms,0,blend_radius_m)
  movel([0.437126, -0.474066, -2.833502, -1.404821, 1.570796, 2.007923],accel_mss,speed_ms,0,blend_radius_m)
  movel([0.438392, -0.474779, -2.833478, -1.404132, 1.570796, 2.009189],accel_mss,speed_ms,0,blend_radius_m)
  movel([0.439295, -0.475904, -2.833441, -1.403044, 1.570796, 2.010091],accel_mss,speed_ms,0,blend_radius_m)
  movel([0.439487, -0.477557, -2.833385, -1.401447, 1.570796, 2.010284],accel_mss,speed_ms,0,blend_radius_m)
  movel([0.439143, -0.479701, -2.833312, -1.399376, 1.570796, 2.009939],accel_mss,speed_ms,0,blend_radius_m)
  movel([0.437530, -0.484736, -2.833133, -1.394520, 1.570796, 2.008326],accel_mss,speed_ms,0,blend_radius_m)
  movel([0.434579, -0.492337, -2.832847, -1.387205, 1.570796, 2.005376],accel_mss,speed_ms,0,blend_radius_m)
  movel([0.431281, -0.500103, -2.832534, -1.379752, 1.570796, 2.002077],accel_mss,speed_ms,0,blend_radius_m)
  movel([0.427645, -0.507997, -2.832194, -1.372198, 1.570796, 1.998441],accel_mss,speed_ms,0,blend_radius_m)
  movel([0.423704, -0.515986, -2.831828, -1.364575, 1.570796, 1.994500],accel_mss,speed_ms,0,blend_radius_m)
  movel([0.419475, -0.524026, -2.831438, -1.356925, 1.570796, 1.990272],accel_mss,speed_ms,0,blend_radius_m)
  movel([0.414991, -0.532081, -2.831023, -1.349285, 1.570796, 1.985787],accel_mss,speed_ms,0,blend_radius_m)
  movel([0.410254, -0.540127, -2.830587, -1.341675, 1.570796, 1.981050],accel_mss,speed_ms,0,blend_radius_m)
  movel([0.405294, -0.548131, -2.830129, -1.334129, 1.570796, 1.976090],accel_mss,speed_ms,0,blend_radius_m)
  movel([0.401988, -0.553148, -2.829830, -1.329410, 1.570796, 1.972784],accel_mss,speed_ms,0,blend_radius_m)
  movel([0.398403, -0.558053, -2.829530, -1.324806, 1.570796, 1.969199],accel_mss,speed_ms,0,blend_radius_m)
  movel([0.394613, -0.562467, -2.829251, -1.320670, 1.570796, 1.965409],accel_mss,speed_ms,0,blend_radius_m)
  movel([0.392667, -0.564361, -2.829130, -1.318898, 1.570796, 1.963463],accel_mss,speed_ms,0,blend_radius_m)
  movel([0.390691, -0.566000, -2.829024, -1.317366, 1.570796, 1.961488],accel_mss,speed_ms,0,blend_radius_m)
  speed_ms = 0.005
  movel([0.390691, -0.560854, -2.822137, -1.329397, 1.570796, 1.961488],accel_mss,speed_ms,0,blend_radius_m)
  speed_ms = 0.040
  movel([0.379771, -0.574577, -2.821211, -1.316601, 1.570796, 1.950568],accel_mss,speed_ms,0,blend_radius_m)
  speed_ms = 0.005
  movel([0.379771, -0.579970, -2.828078, -1.304342, 1.570796, 1.950568],accel_mss,speed_ms,0,blend_radius_m)
  speed_ms = 0.025
  movel([0.379949, -0.581034, -2.828003, -1.303352, 1.570796, 1.950745],accel_mss,speed_ms,0,blend_radius_m)
  movel([0.379468, -0.582647, -2.827888, -1.301854, 1.570796, 1.950264],accel_mss,speed_ms,0,blend_radius_m)
  movel([0.378499, -0.584532, -2.827753, -1.300104, 1.570796, 1.949295],accel_mss,speed_ms,0,blend_radius_m)
  movel([0.377199, -0.586416, -2.827617, -1.298356, 1.570796, 1.947995],accel_mss,speed_ms,0,blend_radius_m)
  movel([0.375432, -0.588327, -2.827477, -1.296585, 1.570796, 1.946228],accel_mss,speed_ms,0,blend_radius_m)
  movel([0.373657, -0.589843, -2.827365, -1.295180, 1.570796, 1.944453],accel_mss,speed_ms,0,blend_radius_m)
  movel([0.371926, -0.591264, -2.827260, -1.293865, 1.570796, 1.942722],accel_mss,speed_ms,0,blend_radius_m)
  movel([0.370313, -0.592885, -2.827139, -1.292365, 1.570796, 1.941109],accel_mss,speed_ms,0,blend_radius_m)
  movel([0.368536, -0.595626, -2.826931, -1.289832, 1.570796, 1.939332],accel_mss,speed_ms,0,blend_radius_m)
  movel([0.367706, -0.597051, -2.826822, -1.288516, 1.570796, 1.938503],accel_mss,speed_ms,0,blend_radius_m)
  movel([0.366616, -0.598563, -2.826706, -1.287120, 1.570796, 1.937412],accel_mss,speed_ms,0,blend_radius_m)
  movel([0.363281, -0.602313, -2.826413, -1.283663, 1.570796, 1.934078],accel_mss,speed_ms,0,blend_radius_m)
  movel([0.359964, -0.605537, -2.826157, -1.280694, 1.570796, 1.930761],accel_mss,speed_ms,0,blend_radius_m)
  movel([0.356635, -0.608317, -2.825934, -1.278139, 1.570796, 1.927431],accel_mss,speed_ms,0,blend_radius_m)
  movel([0.353259, -0.610760, -2.825734, -1.275895, 1.570796, 1.924055],accel_mss,speed_ms,0,blend_radius_m)
  movel([0.355034, -0.609309, -2.825853, -1.277227, 1.570796, 1.925830],accel_mss,speed_ms,0,blend_radius_m)
  movel([0.356757, -0.608140, -2.825948, -1.278301, 1.570796, 1.927553],accel_mss,speed_ms,0,blend_radius_m)
  movel([0.358252, -0.607624, -2.825990, -1.278776, 1.570796, 1.929048],accel_mss,speed_ms,0,blend_radius_m)
  movel([0.359104, -0.608124, -2.825949, -1.278316, 1.570796, 1.929901],accel_mss,speed_ms,0,blend_radius_m)
  movel([0.358949, -0.609664, -2.825824, -1.276901, 1.570796, 1.929745],accel_mss,speed_ms,0,blend_radius_m)
  movel([0.358015, -0.611685, -2.825658, -1.275046, 1.570796, 1.928811],accel_mss,speed_ms,0,blend_radius_m)
  movel([0.356611, -0.613733, -2.825489, -1.273167, 1.570796, 1.927407],accel_mss,speed_ms,0,blend_radius_m)
  movel([0.352353, -0.618606, -2.825079, -1.268704, 1.570796, 1.923149],accel_mss,speed_ms,0,blend_radius_m)
  movel([0.349628, -0.621300, -2.824849, -1.266241, 1.570796, 1.920424],accel_mss,speed_ms,0,blend_radius_m)
  movel([0.346894, -0.623711, -2.824640, -1.264038, 1.570796, 1.917690],accel_mss,speed_ms,0,blend_radius_m)
  movel([0.344176, -0.625813, -2.824456, -1.262120, 1.570796, 1.914972],accel_mss,speed_ms,0,blend_radius_m)
  movel([0.347204, -0.623870, -2.824626, -1.263893, 1.570796, 1.918001],accel_mss,speed_ms,0,blend_radius_m)
  movel([0.350417, -0.621449, -2.824836, -1.266104, 1.570796, 1.921214],accel_mss,speed_ms,0,blend_radius_m)
  movel([0.353558, -0.619146, -2.825033, -1.268210, 1.570796, 1.924354],accel_mss,speed_ms,0,blend_radius_m)
  movel([0.356373, -0.617533, -2.825170, -1.269686, 1.570796, 1.927169],accel_mss,speed_ms,0,blend_radius_m)
  movel([0.357104, -0.617459, -2.825176, -1.269754, 1.570796, 1.927900],accel_mss,speed_ms,0,blend_radius_m)
  movel([0.357042, -0.618082, -2.825124, -1.269184, 1.570796, 1.927838],accel_mss,speed_ms,0,blend_radius_m)
  movel([0.355138, -0.621420, -2.824838, -1.266131, 1.570796, 1.925934],accel_mss,speed_ms,0,blend_radius_m)
  movel([0.353460, -0.623843, -2.824628, -1.263918, 1.570796, 1.924257],accel_mss,speed_ms,0,blend_radius_m)
  movel([0.351629, -0.626168, -2.824425, -1.261797, 1.570796, 1.922426],accel_mss,speed_ms,0,blend_radius_m)
  movel([0.349693, -0.628332, -2.824234, -1.259823, 1.570796, 1.920490],accel_mss,speed_ms,0,blend_radius_m)
  movel([0.350644, -0.627490, -2.824308, -1.260590, 1.570796, 1.921441],accel_mss,speed_ms,0,blend_radius_m)
  movel([0.351670, -0.626851, -2.824365, -1.261173, 1.570796, 1.922466],accel_mss,speed_ms,0,blend_radius_m)
  movel([0.353820, -0.626130, -2.824428, -1.261831, 1.570796, 1.924616],accel_mss,speed_ms,0,blend_radius_m)
  movel([0.355869, -0.626097, -2.824431, -1.261861, 1.570796, 1.926665],accel_mss,speed_ms,0,blend_radius_m)
  movel([0.357562, -0.626666, -2.824381, -1.261342, 1.570796, 1.928358],accel_mss,speed_ms,0,blend_radius_m)
  movel([0.358648, -0.627745, -2.824286, -1.260358, 1.570796, 1.929444],accel_mss,speed_ms,0,blend_radius_m)
  movel([0.358876, -0.629236, -2.824153, -1.259000, 1.570796, 1.929673],accel_mss,speed_ms,0,blend_radius_m)
  movel([0.358591, -0.630105, -2.824075, -1.258209, 1.570796, 1.929388],accel_mss,speed_ms,0,blend_radius_m)
  movel([0.357999, -0.631038, -2.823992, -1.257360, 1.570796, 1.928795],accel_mss,speed_ms,0,blend_radius_m)
  movel([0.357072, -0.632032, -2.823902, -1.256455, 1.570796, 1.927869],accel_mss,speed_ms,0,blend_radius_m)
  movel([0.355773, -0.633068, -2.823808, -1.255513, 1.570796, 1.926569],accel_mss,speed_ms,0,blend_radius_m)
  movel([0.354385, -0.633815, -2.823740, -1.254834, 1.570796, 1.925181],accel_mss,speed_ms,0,blend_radius_m)
  movel([0.349446, -0.634661, -2.823663, -1.254064, 1.570796, 1.920242],accel_mss,speed_ms,0,blend_radius_m)
  movel([0.347504, -0.635123, -2.823621, -1.253645, 1.570796, 1.918301],accel_mss,speed_ms,0,blend_radius_m)
  movel([0.345366, -0.636051, -2.823536, -1.252802, 1.570796, 1.916163],accel_mss,speed_ms,0,blend_radius_m)
  movel([0.341503, -0.638684, -2.823292, -1.250413, 1.570796, 1.912300],accel_mss,speed_ms,0,blend_radius_m)
  movel([0.337576, -0.641615, -2.823018, -1.247756, 1.570796, 1.908372],accel_mss,speed_ms,0,blend_radius_m)
  movel([0.335660, -0.642745, -2.822912, -1.246733, 1.570796, 1.906456],accel_mss,speed_ms,0,blend_radius_m)
  movel([0.333925, -0.643387, -2.822851, -1.246152, 1.570796, 1.904721],accel_mss,speed_ms,0,blend_radius_m)
  movel([0.332602, -0.643348, -2.822854, -1.246186, 1.570796, 1.903398],accel_mss,speed_ms,0,blend_radius_m)
  movel([0.331912, -0.642450, -2.822939, -1.247000, 1.570796, 1.902709],accel_mss,speed_ms,0,blend_radius_m)
  movel([0.333990, -0.639687, -2.823199, -1.249503, 1.570796, 1.904787],accel_mss,speed_ms,0,blend_radius_m)
  movel([0.336211, -0.637050, -2.823444, -1.251895, 1.570796, 1.907007],accel_mss,speed_ms,0,blend_radius_m)
  speed_ms = 0.005
  movel([0.336211, -0.630701, -2.816672, -1.265016, 1.570796, 1.907007],accel_mss,speed_ms,0,blend_radius_m)
  speed_ms = 0.040
  movel([0.351549, -0.640243, -2.815776, -1.256370, 1.570796, 1.922345],accel_mss,speed_ms,0,blend_radius_m)
  speed_ms = 0.005
  movel([0.351549, -0.646746, -2.822530, -1.243114, 1.570796, 1.922345],accel_mss,speed_ms,0,blend_radius_m)
  speed_ms = 0.025
  movel([0.353017, -0.644776, -2.822719, -1.244895, 1.570796, 1.923813],accel_mss,speed_ms,0,blend_radius_m)
  movel([0.354736, -0.643268, -2.822862, -1.246259, 1.570796, 1.925532],accel_mss,speed_ms,0,blend_radius_m)
  movel([0.356426, -0.642349, -2.822949, -1.247091, 1.570796, 1.927223],accel_mss,speed_ms,0,blend_radius_m)
  movel([0.357799, -0.642160, -2.822967, -1.247262, 1.570796, 1.928595],accel_mss,speed_ms,0,blend_radius_m)
  movel([0.358713, -0.642649, -2.822921, -1.246819, 1.570796, 1.929509],accel_mss,speed_ms,0,blend_radius_m)
  movel([0.359289, -0.643571, -2.822833, -1.245985, 1.570796, 1.930085],accel_mss,speed_ms,0,blend_radius_m)
  movel([0.359851, -0.646096, -2.822592, -1.243701, 1.570796, 1.930648],accel_mss,speed_ms,0,blend_radius_m)
  movel([0.361230, -0.643691, -2.822822, -1.245876, 1.570796, 1.932027],accel_mss,speed_ms,0,blend_radius_m)
  movel([0.362162, -0.641381, -2.823040, -1.247968, 1.570796, 1.932958],accel_mss,speed_ms,0,blend_radius_m)
  movel([0.362570, -0.639367, -2.823229, -1.249793, 1.570796, 1.933367],accel_mss,speed_ms,0,blend_radius_m)
  movel([0.362409, -0.637813, -2.823373, -1.251203, 1.570796, 1.933205],accel_mss,speed_ms,0,blend_radius_m)
  movel([0.363247, -0.638243, -2.823333, -1.250813, 1.570796, 1.934044],accel_mss,speed_ms,0,blend_radius_m)
  movel([0.363803, -0.639012, -2.823262, -1.250115, 1.570796, 1.934599],accel_mss,speed_ms,0,blend_radius_m)
  movel([0.364218, -0.641334, -2.823045, -1.248010, 1.570796, 1.935014],accel_mss,speed_ms,0,blend_radius_m)
  movel([0.363986, -0.644333, -2.822761, -1.245295, 1.570796, 1.934783],accel_mss,speed_ms,0,blend_radius_m)
  movel([0.363403, -0.647600, -2.822447, -1.242342, 1.570796, 1.934200],accel_mss,speed_ms,0,blend_radius_m)
  movel([0.362304, -0.651413, -2.822076, -1.238900, 1.570796, 1.933101],accel_mss,speed_ms,0,blend_radius_m)
  movel([0.360800, -0.655221, -2.821700, -1.235468, 1.570796, 1.931596],accel_mss,speed_ms,0,blend_radius_m)
  movel([0.359255, -0.658978, -2.821322, -1.232089, 1.570796, 1.930051],accel_mss,speed_ms,0,blend_radius_m)
  movel([0.358028, -0.662650, -2.820948, -1.228791, 1.570796, 1.928824],accel_mss,speed_ms,0,blend_radius_m)
  movel([0.357067, -0.661034, -2.821113, -1.230242, 1.570796, 1.927863],accel_mss,speed_ms,0,blend_radius_m)
  movel([0.355532, -0.660158, -2.821203, -1.231029, 1.570796, 1.926329],accel_mss,speed_ms,0,blend_radius_m)
  movel([0.353464, -0.660097, -2.821209, -1.231083, 1.570796, 1.924261],accel_mss,speed_ms,0,blend_radius_m)
  movel([0.350894, -0.660931, -2.821124, -1.230334, 1.570796, 1.921690],accel_mss,speed_ms,0,blend_radius_m)
  speed_ms = 0.005
  movel([0.350894, -0.654209, -2.814398, -1.243782, 1.570796, 1.921690],accel_mss,speed_ms,0,blend_radius_m)
  speed_ms = 0.040
  movel([0.352138, -0.663792, -2.813406, -1.235191, 1.570796, 1.922935],accel_mss,speed_ms,0,blend_radius_m)
  speed_ms = 0.005
  movel([0.352138, -0.670661, -2.820112, -1.221617, 1.570796, 1.922935],accel_mss,speed_ms,0,blend_radius_m)
  speed_ms = 0.025
  movel([0.351964, -0.674802, -2.819669, -1.217918, 1.570796, 1.922760],accel_mss,speed_ms,0,blend_radius_m)
  movel([0.352428, -0.678371, -2.819281, -1.214737, 1.570796, 1.923224],accel_mss,speed_ms,0,blend_radius_m)
  movel([0.353764, -0.680933, -2.819000, -1.212456, 1.570796, 1.924560],accel_mss,speed_ms,0,blend_radius_m)
  movel([0.354836, -0.681702, -2.818915, -1.211772, 1.570796, 1.925632],accel_mss,speed_ms,0,blend_radius_m)
  movel([0.356219, -0.682058, -2.818875, -1.211455, 1.570796, 1.927016],accel_mss,speed_ms,0,blend_radius_m)
  movel([0.358558, -0.681811, -2.818903, -1.211675, 1.570796, 1.929355],accel_mss,speed_ms,0,blend_radius_m)
  movel([0.361206, -0.680840, -2.819010, -1.212539, 1.570796, 1.932002],accel_mss,speed_ms,0,blend_radius_m)
  movel([0.364101, -0.679308, -2.819179, -1.213902, 1.570796, 1.934897],accel_mss,speed_ms,0,blend_radius_m)
  movel([0.367174, -0.677385, -2.819389, -1.215615, 1.570796, 1.937971],accel_mss,speed_ms,0,blend_radius_m)
  movel([0.373586, -0.673021, -2.819860, -1.219507, 1.570796, 1.944382],accel_mss,speed_ms,0,blend_radius_m)
  movel([0.379870, -0.669113, -2.820275, -1.223000, 1.570796, 1.950666],accel_mss,speed_ms,0,blend_radius_m)
  movel([0.383258, -0.667573, -2.820437, -1.224379, 1.570796, 1.954054],accel_mss,speed_ms,0,blend_radius_m)
  movel([0.386363, -0.666706, -2.820528, -1.225155, 1.570796, 1.957160],accel_mss,speed_ms,0,blend_radius_m)
  movel([0.389136, -0.666499, -2.820549, -1.225341, 1.570796, 1.959932],accel_mss,speed_ms,0,blend_radius_m)
  movel([0.391521, -0.666944, -2.820503, -1.224942, 1.570796, 1.962317],accel_mss,speed_ms,0,blend_radius_m)
  movel([0.393479, -0.668012, -2.820391, -1.223986, 1.570796, 1.964275],accel_mss,speed_ms,0,blend_radius_m)
  movel([0.394959, -0.669692, -2.820214, -1.222483, 1.570796, 1.965755],accel_mss,speed_ms,0,blend_radius_m)
  movel([0.395914, -0.671962, -2.819973, -1.220453, 1.570796, 1.966710],accel_mss,speed_ms,0,blend_radius_m)
  movel([0.396312, -0.674790, -2.819670, -1.217929, 1.570796, 1.967108],accel_mss,speed_ms,0,blend_radius_m)
  speed_ms = 0.005
  movel([0.396312, -0.667859, -2.812973, -1.231557, 1.570796, 1.967108],accel_mss,speed_ms,0,blend_radius_m)
  speed_ms = 0.040
  movel([0.345905, -0.635640, -2.816213, -1.260537, 1.570796, 1.916701],accel_mss,speed_ms,0,blend_radius_m)
  speed_ms = 0.005
  movel([0.345905, -0.642068, -2.822975, -1.247345, 1.570796, 1.916701],accel_mss,speed_ms,0,blend_radius_m)
  speed_ms = 0.025
  movel([0.347293, -0.642385, -2.822946, -1.247058, 1.570796, 1.918089],accel_mss,speed_ms,0,blend_radius_m)
  movel([0.348210, -0.643311, -2.822858, -1.246220, 1.570796, 1.919007],accel_mss,speed_ms,0,blend_radius_m)
  movel([0.348304, -0.644184, -2.822775, -1.245430, 1.570796, 1.919100],accel_mss,speed_ms,0,blend_radius_m)
  movel([0.348070, -0.645320, -2.822667, -1.244402, 1.570796, 1.918866],accel_mss,speed_ms,0,blend_radius_m)
  movel([0.347517, -0.646595, -2.822544, -1.243249, 1.570796, 1.918313],accel_mss,speed_ms,0,blend_radius_m)
  movel([0.346644, -0.647884, -2.822420, -1.242085, 1.570796, 1.917440],accel_mss,speed_ms,0,blend_radius_m)
  movel([0.344727, -0.650018, -2.822213, -1.240158, 1.570796, 1.915523],accel_mss,speed_ms,0,blend_radius_m)
  movel([0.343988, -0.651235, -2.822094, -1.239060, 1.570796, 1.914784],accel_mss,speed_ms,0,blend_radius_m)
  movel([0.343592, -0.652382, -2.821981, -1.238026, 1.570796, 1.914388],accel_mss,speed_ms,0,blend_radius_m)
  movel([0.343551, -0.654276, -2.821794, -1.236320, 1.570796, 1.914347],accel_mss,speed_ms,0,blend_radius_m)
  movel([0.344108, -0.655922, -2.821630, -1.234837, 1.570796, 1.914905],accel_mss,speed_ms,0,blend_radius_m)
  movel([0.345022, -0.657166, -2.821505, -1.233718, 1.570796, 1.915818],accel_mss,speed_ms,0,blend_radius_m)
  movel([0.346266, -0.658001, -2.821421, -1.232967, 1.570796, 1.917062],accel_mss,speed_ms,0,blend_radius_m)
  movel([0.347814, -0.658397, -2.821381, -1.232611, 1.570796, 1.918611],accel_mss,speed_ms,0,blend_radius_m)
  movel([0.346143, -0.661118, -2.821105, -1.230166, 1.570796, 1.916940],accel_mss,speed_ms,0,blend_radius_m)
  movel([0.344813, -0.663764, -2.820833, -1.227792, 1.570796, 1.915609],accel_mss,speed_ms,0,blend_radius_m)
  movel([0.343783, -0.666330, -2.820567, -1.225492, 1.570796, 1.914580],accel_mss,speed_ms,0,blend_radius_m)
  movel([0.343015, -0.668806, -2.820308, -1.223275, 1.570796, 1.913812],accel_mss,speed_ms,0,blend_radius_m)
  movel([0.342123, -0.673455, -2.819814, -1.219120, 1.570796, 1.912920],accel_mss,speed_ms,0,blend_radius_m)
  movel([0.341863, -0.677637, -2.819361, -1.215390, 1.570796, 1.912659],accel_mss,speed_ms,0,blend_radius_m)
  movel([0.341691, -0.681612, -2.818925, -1.211852, 1.570796, 1.912487],accel_mss,speed_ms,0,blend_radius_m)
  movel([0.341301, -0.683792, -2.818683, -1.209914, 1.570796, 1.912097],accel_mss,speed_ms,0,blend_radius_m)
  movel([0.340520, -0.686192, -2.818414, -1.207783, 1.570796, 1.911316],accel_mss,speed_ms,0,blend_radius_m)
  movel([0.339172, -0.688831, -2.818115, -1.205443, 1.570796, 1.909969],accel_mss,speed_ms,0,blend_radius_m)
  movel([0.337350, -0.691417, -2.817819, -1.203153, 1.570796, 1.908147],accel_mss,speed_ms,0,blend_radius_m)
  movel([0.335304, -0.693545, -2.817574, -1.201270, 1.570796, 1.906101],accel_mss,speed_ms,0,blend_radius_m)
  movel([0.333296, -0.694803, -2.817428, -1.200158, 1.570796, 1.904092],accel_mss,speed_ms,0,blend_radius_m)
  movel([0.333851, -0.696131, -2.817273, -1.198985, 1.570796, 1.904647],accel_mss,speed_ms,0,blend_radius_m)
  movel([0.334133, -0.699579, -2.816867, -1.195942, 1.570796, 1.904930],accel_mss,speed_ms,0,blend_radius_m)
  movel([0.333871, -0.701631, -2.816623, -1.194134, 1.570796, 1.904667],accel_mss,speed_ms,0,blend_radius_m)
  movel([0.332594, -0.706194, -2.816074, -1.190120, 1.570796, 1.903390],accel_mss,speed_ms,0,blend_radius_m)
  movel([0.331591, -0.708632, -2.815777, -1.187979, 1.570796, 1.902387],accel_mss,speed_ms,0,blend_radius_m)
  movel([0.330351, -0.711135, -2.815470, -1.185785, 1.570796, 1.901147],accel_mss,speed_ms,0,blend_radius_m)
  speed_ms = 0.005
  movel([0.330351, -0.703686, -2.808854, -1.199849, 1.570796, 1.901147],accel_mss,speed_ms,0,blend_radius_m)
  speed_ms = 0.040
  movel([0.320831, -0.707801, -2.808345, -1.196243, 1.570796, 1.891628],accel_mss,speed_ms,0,blend_radius_m)
  speed_ms = 0.005
  movel([0.320831, -0.715307, -2.814951, -1.182132, 1.570796, 1.891628],accel_mss,speed_ms,0,blend_radius_m)
  speed_ms = 0.025
  movel([0.323413, -0.732368, -2.812746, -1.167275, 1.570796, 1.894209],accel_mss,speed_ms,0,blend_radius_m)
  movel([0.323461, -0.734669, -2.812439, -1.165281, 1.570796, 1.894258],accel_mss,speed_ms,0,blend_radius_m)
  movel([0.323113, -0.736017, -2.812258, -1.164114, 1.570796, 1.893909],accel_mss,speed_ms,0,blend_radius_m)
  movel([0.322352, -0.737486, -2.812059, -1.162844, 1.570796, 1.893148],accel_mss,speed_ms,0,blend_radius_m)
  movel([0.320056, -0.740590, -2.811637, -1.160163, 1.570796, 1.890852],accel_mss,speed_ms,0,blend_radius_m)
  movel([0.319501, -0.742123, -2.811426, -1.158840, 1.570796, 1.890297],accel_mss,speed_ms,0,blend_radius_m)
  movel([0.319482, -0.743376, -2.811254, -1.157760, 1.570796, 1.890279],accel_mss,speed_ms,0,blend_radius_m)
  movel([0.320112, -0.744880, -2.811045, -1.156464, 1.570796, 1.890908],accel_mss,speed_ms,0,blend_radius_m)
  movel([0.321291, -0.745853, -2.810910, -1.155626, 1.570796, 1.892088],accel_mss,speed_ms,0,blend_radius_m)
  movel([0.323990, -0.747265, -2.810713, -1.154411, 1.570796, 1.894786],accel_mss,speed_ms,0,blend_radius_m)
  movel([0.325329, -0.748755, -2.810504, -1.153130, 1.570796, 1.896125],accel_mss,speed_ms,0,blend_radius_m)
  movel([0.326698, -0.751442, -2.810124, -1.150823, 1.570796, 1.897494],accel_mss,speed_ms,0,blend_radius_m)
  movel([0.326968, -0.752971, -2.809906, -1.149512, 1.570796, 1.897764],accel_mss,speed_ms,0,blend_radius_m)
  movel([0.326754, -0.754472, -2.809692, -1.148226, 1.570796, 1.897550],accel_mss,speed_ms,0,blend_radius_m)
  movel([0.326410, -0.755177, -2.809590, -1.147622, 1.570796, 1.897207],accel_mss,speed_ms,0,blend_radius_m)
  movel([0.325881, -0.755833, -2.809496, -1.147060, 1.570796, 1.896678],accel_mss,speed_ms,0,blend_radius_m)
  movel([0.324184, -0.756962, -2.809333, -1.146094, 1.570796, 1.894981],accel_mss,speed_ms,0,blend_radius_m)
  movel([0.324146, -0.758452, -2.809117, -1.144820, 1.570796, 1.894943],accel_mss,speed_ms,0,blend_radius_m)
  movel([0.324547, -0.759800, -2.808921, -1.143668, 1.570796, 1.895344],accel_mss,speed_ms,0,blend_radius_m)
  movel([0.326252, -0.762067, -2.808589, -1.141733, 1.570796, 1.897049],accel_mss,speed_ms,0,blend_radius_m)
  movel([0.330428, -0.764958, -2.808162, -1.139270, 1.570796, 1.901225],accel_mss,speed_ms,0,blend_radius_m)
  movel([0.332973, -0.765749, -2.808044, -1.138596, 1.570796, 1.903769],accel_mss,speed_ms,0,blend_radius_m)
  movel([0.335888, -0.766200, -2.807977, -1.138212, 1.570796, 1.906684],accel_mss,speed_ms,0,blend_radius_m)
  movel([0.338411, -0.767130, -2.807838, -1.137421, 1.570796, 1.909207],accel_mss,speed_ms,0,blend_radius_m)
  movel([0.339288, -0.768024, -2.807704, -1.136661, 1.570796, 1.910085],accel_mss,speed_ms,0,blend_radius_m)
  movel([0.339784, -0.769337, -2.807507, -1.135545, 1.570796, 1.910580],accel_mss,speed_ms,0,blend_radius_m)
  movel([0.339779, -0.770249, -2.807370, -1.134770, 1.570796, 1.910575],accel_mss,speed_ms,0,blend_radius_m)
  movel([0.339496, -0.771333, -2.807206, -1.133850, 1.570796, 1.910293],accel_mss,speed_ms,0,blend_radius_m)
  movel([0.338944, -0.772395, -2.807044, -1.132950, 1.570796, 1.909740],accel_mss,speed_ms,0,blend_radius_m)
  movel([0.338115, -0.773237, -2.806916, -1.132236, 1.570796, 1.908911],accel_mss,speed_ms,0,blend_radius_m)
  movel([0.336844, -0.773572, -2.806865, -1.131952, 1.570796, 1.907640],accel_mss,speed_ms,0,blend_radius_m)
  movel([0.331845, -0.772888, -2.806969, -1.132531, 1.570796, 1.902641],accel_mss,speed_ms,0,blend_radius_m)
  movel([0.327463, -0.771244, -2.807219, -1.133926, 1.570796, 1.898259],accel_mss,speed_ms,0,blend_radius_m)
  movel([0.326911, -0.772441, -2.807037, -1.132910, 1.570796, 1.897708],accel_mss,speed_ms,0,blend_radius_m)
  movel([0.326609, -0.773547, -2.806869, -1.131973, 1.570796, 1.897405],accel_mss,speed_ms,0,blend_radius_m)
  movel([0.326653, -0.775494, -2.806571, -1.130324, 1.570796, 1.897450],accel_mss,speed_ms,0,blend_radius_m)
  movel([0.327394, -0.777112, -2.806322, -1.128955, 1.570796, 1.898190],accel_mss,speed_ms,0,blend_radius_m)
  movel([0.328616, -0.778453, -2.806114, -1.127822, 1.570796, 1.899412],accel_mss,speed_ms,0,blend_radius_m)
  movel([0.331744, -0.780391, -2.805813, -1.126185, 1.570796, 1.902540],accel_mss,speed_ms,0,blend_radius_m)
  movel([0.334451, -0.781554, -2.805631, -1.125204, 1.570796, 1.905247],accel_mss,speed_ms,0,blend_radius_m)
  movel([0.335324, -0.782159, -2.805537, -1.124694, 1.570796, 1.906121],accel_mss,speed_ms,0,blend_radius_m)
  movel([0.335511, -0.782701, -2.805451, -1.124237, 1.570796, 1.906307],accel_mss,speed_ms,0,blend_radius_m)
  movel([0.335387, -0.783482, -2.805329, -1.123579, 1.570796, 1.906183],accel_mss,speed_ms,0,blend_radius_m)
  movel([0.334923, -0.784452, -2.805175, -1.122761, 1.570796, 1.905720],accel_mss,speed_ms,0,blend_radius_m)
  movel([0.334354, -0.785155, -2.805064, -1.122170, 1.570796, 1.905150],accel_mss,speed_ms,0,blend_radius_m)
  movel([0.333034, -0.786032, -2.804925, -1.121432, 1.570796, 1.903831],accel_mss,speed_ms,0,blend_radius_m)
  movel([0.331203, -0.787058, -2.804762, -1.120569, 1.570796, 1.901999],accel_mss,speed_ms,0,blend_radius_m)
  movel([0.330790, -0.787594, -2.804677, -1.120118, 1.570796, 1.901586],accel_mss,speed_ms,0,blend_radius_m)
  movel([0.330501, -0.788396, -2.804549, -1.119445, 1.570796, 1.901297],accel_mss,speed_ms,0,blend_radius_m)
  movel([0.330491, -0.789128, -2.804431, -1.118830, 1.570796, 1.901287],accel_mss,speed_ms,0,blend_radius_m)
  movel([0.331058, -0.790375, -2.804231, -1.117783, 1.570796, 1.901854],accel_mss,speed_ms,0,blend_radius_m)
  movel([0.332754, -0.792042, -2.803962, -1.116385, 1.570796, 1.903551],accel_mss,speed_ms,0,blend_radius_m)
  movel([0.340812, -0.798016, -2.802986, -1.111386, 1.570796, 1.911608],accel_mss,speed_ms,0,blend_radius_m)
  movel([0.341451, -0.798829, -2.802852, -1.110708, 1.570796, 1.912247],accel_mss,speed_ms,0,blend_radius_m)
  movel([0.341793, -0.799946, -2.802667, -1.109776, 1.570796, 1.912589],accel_mss,speed_ms,0,blend_radius_m)
  movel([0.341637, -0.801326, -2.802438, -1.108625, 1.570796, 1.912433],accel_mss,speed_ms,0,blend_radius_m)
  movel([0.340781, -0.802917, -2.802172, -1.107300, 1.570796, 1.911578],accel_mss,speed_ms,0,blend_radius_m)
  movel([0.339541, -0.804143, -2.801966, -1.106280, 1.570796, 1.910338],accel_mss,speed_ms,0,blend_radius_m)
  movel([0.338270, -0.804764, -2.801862, -1.105763, 1.570796, 1.909067],accel_mss,speed_ms,0,blend_radius_m)
